                       3: //System 3
                           IF #_id_decoded_OP[#i].Device_Type = 30 THEN //VTD
                               "Screen_DB".OrderProcessing[#i] := CONCAT(IN1 := "System_DB_3".OrderTable[1].Device, IN2 := ' To LEVEL ', IN3 := #Level_Strg);
                           ELSIF #_id_decoded_OP[#i].Device_Type = 10 THEN //CNV1
                               "Screen_DB".OrderProcessing[#i] := CONCAT(IN1 := "System_DB_3".OrderTable[1].Device, IN2 := ' To CNV 1 LEVEL ', IN3 := #Level_Strg);
                           ELSIF #_id_decoded_OP[#i].Device_Type = 11 THEN //CNV2
                               "Screen_DB".OrderProcessing[#i] := CONCAT(IN1 := "System_DB_3".OrderTable[1].Device, IN2 := ' To CNV 2 LEVEL ', IN3 := #Level_Strg);
                           ELSIF #_id_decoded_OP[#i].Device_Type = 12 THEN //ECONVEYOR
                               "Screen_DB".OrderProcessing[#i] := CONCAT(IN1 := "System_DB_3".OrderTable[1].Device, IN2 := ' To ECONV LEVEL ', IN3 := #Level_Strg);
                           END_IF;

                       4: //System 4
                           IF #_id_decoded_OP[#i].Device_Type = 30 THEN //VTD
                               "Screen_DB".OrderProcessing[#i] := CONCAT(IN1 := "System_DB_4".OrderTable[1].Device, IN2 := ' To LEVEL ', IN3 := #Level_Strg);
                           ELSIF #_id_decoded_OP[#i].Device_Type = 10 THEN //CNV1
                               "Screen_DB".OrderProcessing[#i] := CONCAT(IN1 := "System_DB_4".OrderTable[1].Device, IN2 := ' To CNV 1 LEVEL ', IN3 := #Level_Strg);
                           ELSIF #_id_decoded_OP[#i].Device_Type = 11 THEN //CNV2
                               "Screen_DB".OrderProcessing[#i] := CONCAT(IN1 := "System_DB_4".OrderTable[1].Device, IN2 := ' To CNV 2 LEVEL ', IN3 := #Level_Strg);
                           ELSIF #_id_decoded_OP[#i].Device_Type = 12 THEN //ECONVEYOR
                               "Screen_DB".OrderProcessing[#i] := CONCAT(IN1 := "System_DB_4".OrderTable[1].Device, IN2 := ' To ECONV LEVEL ', IN3 := #Level_Strg);
                           END_IF;

                       5: //System 5
                           IF #_id_decoded_OP[#i].Device_Type = 30 THEN //VTD
                               "Screen_DB".OrderProcessing[#i] := CONCAT(IN1 := "System_DB_5".OrderTable[1].Device, IN2 := ' To LEVEL ', IN3 := #Level_Strg);
                           ELSIF #_id_decoded_OP[#i].Device_Type = 10 THEN //CNV1
                               "Screen_DB".OrderProcessing[#i] := CONCAT(IN1 := "System_DB_5".OrderTable[1].Device, IN2 := ' To CNV 1 LEVEL ', IN3 := #Level_Strg);
                           ELSIF #_id_decoded_OP[#i].Device_Type = 11 THEN //CNV2
                               "Screen_DB".OrderProcessing[#i] := CONCAT(IN1 := "System_DB_5".OrderTable[1].Device, IN2 := ' To CNV 2 LEVEL ', IN3 := #Level_Strg);
                           ELSIF #_id_decoded_OP[#i].Device_Type = 12 THEN //ECONVEYOR
                               "Screen_DB".OrderProcessing[#i] := CONCAT(IN1 := "System_DB_5".OrderTable[1].Device, IN2 := ' To ECONV LEVEL ', IN3 := #Level_Strg);
                           END_IF;
                   END_CASE;
               END_IF;
               END_FOR;

       END_REGION

       //empty background
       IF "System_DB_1".Error OR "System_DB_2".Error OR "System_DB_3".Error OR "System_DB_4".Error OR "System_DB_5".Error OR
           "Error_Word_1" <> 0 OR
           "Errors_Profinet_1" <> 0 OR
           "Errors_Profinet_2" <> 0 OR
           "Errors_Profinet_3" <> 0 OR
           "Errors_Profinet_4" <> 0 OR
           "Errors_Profinet_5" <> 0 OR
           "Errors_Profinet_6" <> 0 OR
           "Errors_Profinet_7" <> 0 OR
           "Errors_Profinet_8" <> 0 OR
           "Errors_Profinet_9" <> 0 OR
           "Errors_Profinet_10".%X0 OR
           "Errors_Profinet_10".%X1 OR
           "Errors_Profinet_10".%X2 OR
           "Errors_Profinet_10".%X3 OR
           "Errors_Profinet_10".%X4 OR
           "Errors_Profinet_10".%X5 OR
           "Errors_Profinet_10".%X6 OR
           "Errors_Profinet_10".%X7 OR
           "Errors_Profinet_10".%X8 OR
           "Errors_Profinet_10".%X9 OR
           "Errors_Profinet_10".%X10 OR
           "Errors_Profinet_10".%X11 OR
           "Errors_Profinet_10".%X12 OR
           "Errors_Profinet_10".%X13 OR
           "Errors_Profinet_11" <> 0 OR
           "Erros_Supply_Feedback_1" <> 0 OR
           "Erros_Supply_Feedback_2" <> 0 OR
           "Erros_Supply_Feedback_3" <> 0 OR
           "Erros_Supply_Feedback_4" <> 0 OR
           "Erros_Supply_Feedback_5" <> 0 OR
           "Erros_Supply_Feedback_6" <> 0 OR
           "Erros_Supply_Feedback_7" <> 0 OR
           "Sick Lector_Error code 1" <> 0 OR
           "Sick Lector_Error code 2" <> 0 OR
           "Sick Lector_Error code 3" <> 0 OR
           "Sick Lector_Error code 4" <> 0 OR
           "Sick Lector_Error code 5" <> 0 OR
           "Linear Encoder_Device Errors 1" <> 0 OR
           "Linear Encoder_Device Errors 2" <> 0 OR
           "Linear Encoder_Device Errors 3" <> 0 OR
           "Linear Encoder_Device Errors 4" <> 0 OR
           "Linear Encoder_Device Errors 5" <> 0 OR
           "Estop_Error_Word_1" <> 0 OR
           "Estop_Error_Word_2" <> 0 OR
           "Estop_Error_Word_3" <> 0 OR
           "Estop_Error_Word_4" <> 0 OR
           "Estop_Error_Word_5" <> 0 OR
           "Estop_Error_Word_6" <> 0 OR
           "Errors_Word_LightGuard_1" <> 0
       THEN
           "Screen_DB".EmptyTemplate_Background := 1;
       ELSE
           "Screen_DB".EmptyTemplate_Background := 0;
       END_IF;    //e

       // //main background - DEVICES
       // IF "HMI_DB".ScreenNo_Main = 1 AND "VTD_System_Selected_HMI" <> 0 THEN //VTD SCREEN
       //     IF "Control_DB".VTD_Sys["VTD_System_Selected_HMI"]."Error" THEN
       //         "Screen_DB".MainTemplate_Background := 1;
       //     ELSE
       //         "Screen_DB".MainTemplate_Background := 0;
       //     END_IF;
       // ELSIF "HMI_DB".ScreenNo_Main = 2 AND "CNV_System_Selected" <> 0 AND "CNV2_Selected" <> 0 AND "CNV_Level_Selected" <> 0 THEN //CONVEYOR SCREEN
       //     IF "CNV2_Selected" = 1 AND ("Control_DB".LCnv_Sys["CNV_System_Selected"].Cnv_Level["CNV_Level_Selected"].Cnv1.Error OR
       //         "Control_DB".ECnv_Sys["CNV_System_Selected"].Error) THEN
       //         "Screen_DB".MainTemplate_Background := 1;
       //     ELSIF "CNV2_Selected" = 2 AND ("Control_DB".LCnv_Sys["CNV_System_Selected"].Cnv_Level["CNV_Level_Selected"].Cnv2.Error OR
       //         "Control_DB".ECnv_Sys["CNV_System_Selected"].Error) THEN
       //         "Screen_DB".MainTemplate_Background := 1;
       //     ELSE
       //         "Screen_DB".MainTemplate_Background := 0;
       //     END_IF;
       // ELSE
       //     "Screen_DB".MainTemplate_Background := 0;
       // END_IF;
   END_REGION;

   REGION SHUTTLES
       IF "Screen_DB".Shuttle_Select >= 1 AND "Screen_DB".Shuttle_Select <= "Settings_DB".System.Shuttle_Count THEN
           CASE "Screen_DB".Shuttle_Select OF
               1:
                   "Screen_DB".Shuttle := "Shuttle_MQTT_DB".Shuttle_MQTT[1].Message.Shuttle_Status;
               2:
                   "Screen_DB".Shuttle := "Shuttle_MQTT_DB".Shuttle_MQTT[2].Message.Shuttle_Status;
               3:
                   "Screen_DB".Shuttle := "Shuttle_MQTT_DB".Shuttle_MQTT[3].Message.Shuttle_Status;
               4:
                   "Screen_DB".Shuttle := "Shuttle_MQTT_DB".Shuttle_MQTT[4].Message.Shuttle_Status;
               5:
                   "Screen_DB".Shuttle := "Shuttle_MQTT_DB".Shuttle_MQTT[5].Message.Shuttle_Status;
               6:
                   "Screen_DB".Shuttle := "Shuttle_MQTT_DB".Shuttle_MQTT[6].Message.Shuttle_Status;
               7:
                   "Screen_DB".Shuttle := "Shuttle_MQTT_DB".Shuttle_MQTT[7].Message.Shuttle_Status;
               8:
                   "Screen_DB".Shuttle := "Shuttle_MQTT_DB".Shuttle_MQTT[8].Message.Shuttle_Status;
               9:
                   "Screen_DB".Shuttle := "Shuttle_MQTT_DB".Shuttle_MQTT[9].Message.Shuttle_Status;
               10:
                   "Screen_DB".Shuttle := "Shuttle_MQTT_DB".Shuttle_MQTT[10].Message.Shuttle_Status;
               11:
                   "Screen_DB".Shuttle := "Shuttle_MQTT_DB".Shuttle_MQTT[11].Message.Shuttle_Status;
               12:
                   "Screen_DB".Shuttle := "Shuttle_MQTT_DB".Shuttle_MQTT[12].Message.Shuttle_Status;
               13:
                   "Screen_DB".Shuttle := "Shuttle_MQTT_DB".Shuttle_MQTT[13].Message.Shuttle_Status;
               14:
                   "Screen_DB".Shuttle := "Shuttle_MQTT_DB".Shuttle_MQTT[14].Message.Shuttle_Status;
               15:
                   "Screen_DB".Shuttle := "Shuttle_MQTT_DB".Shuttle_MQTT[15].Message.Shuttle_Status;
               16:
                   "Screen_DB".Shuttle := "Shuttle_MQTT_DB".Shuttle_MQTT[16].Message.Shuttle_Status;
               17:
                   "Screen_DB".Shuttle := "Shuttle_MQTT_DB".Shuttle_MQTT[17].Message.Shuttle_Status;
               18:
                   "Screen_DB".Shuttle := "Shuttle_MQTT_DB".Shuttle_MQTT[18].Message.Shuttle_Status;
               19:
                   "Screen_DB".Shuttle := "Shuttle_MQTT_DB".Shuttle_MQTT[19].Message.Shuttle_Status;
               20:
                   "Screen_DB".Shuttle := "Shuttle_MQTT_DB".Shuttle_MQTT[20].Message.Shuttle_Status;
               21:
                   "Screen_DB".Shuttle := "Shuttle_MQTT_DB".Shuttle_MQTT[21].Message.Shuttle_Status;
               22:
                   "Screen_DB".Shuttle := "Shuttle_MQTT_DB".Shuttle_MQTT[22].Message.Shuttle_Status;
               23:
                   "Screen_DB".Shuttle := "Shuttle_MQTT_DB".Shuttle_MQTT[23].Message.Shuttle_Status;
               // 24:
               //     "Screen_DB".Shuttle := "Shuttle_MQTT_DB".Shuttle_MQTT[24].Message.Shuttle_Status;
           END_CASE;
       END_IF;

       //E-STOP
       IF "Charge_Shuttle_Commands" THEN
           CASE "Shuttle_Level_Selected" OF
               1:
                   "Shuttle_Level_EStop" := "L1_Estop";
               2:
                   "Shuttle_Level_EStop" := "L2_Estop";
               3:
                   "Shuttle_Level_EStop" := "L3_Estop";
               4:
                   "Shuttle_Level_EStop" := "L4_Estop";
               5:
                   "Shuttle_Level_EStop" := "L5_Estop";
               6:
                   "Shuttle_Level_EStop" := "L6_Estop";
               7:
                   "Shuttle_Level_EStop" := "L7_Estop";
               8:
                   "Shuttle_Level_EStop" := "L8_Estop";
           END_CASE;
       ELSE
           CASE "Shuttle_Level_Selected" OF
               1:
                   "L1_Estop" := "Shuttle_Level_EStop";
               2:
                   "L2_Estop" := "Shuttle_Level_EStop";
               3:
                   "L3_Estop" := "Shuttle_Level_EStop";
               4:
                   "L4_Estop" := "Shuttle_Level_EStop";
               5:
                   "L5_Estop" := "Shuttle_Level_EStop";
               6:
                   "L6_Estop" := "Shuttle_Level_EStop";
               7:
                   "L7_Estop" := "Shuttle_Level_EStop";
               8:
                   "L8_Estop" := "Shuttle_Level_EStop";
           END_CASE;
       END_IF;
   END_REGION

   REGION ORDER TABLE
       //CHARGE OT DATA
       IF "Screen_DB".Charge_OT THEN
           CASE "Main_OrderTable_Selected" OF
               1:
                   "OT_Charge_Commands"("Auto_Test_1_DB");
               2:
                   "OT_Charge_Commands"("Auto_Test_2_DB");
               3:
                   "OT_Charge_Commands"("Auto_Test_3_DB");
               4:
                   "OT_Charge_Commands_1"("Auto_Test_4_DB");
               5:
                   "OT_Charge_Commands_1"("Auto_Test_5_DB");
           END_CASE;
           "T_Charge_OT".TON(IN := TRUE,
                             PT := T#1000ms);
           IF "T_Charge_OT".Q THEN
               "T_Charge_OT".TON(IN := FALSE,
                                 PT := T#0ms);
               "Screen_DB".Charge_OT := FALSE;
           END_IF;
       END_IF;

       IF NOT "Screen_DB".Charge_OT THEN
           "T_Charge_OT".TON(IN := FALSE,
                             PT := T#0ms);

           CASE "Main_OrderTable_Selected" OF
               1:
                   "Clear_OT(1)" := "Clear_OT";
                   "FC_Orders"(Sys := 1,
                               System := "System_DB_1",
                               Auto_Test := "Auto_Test_1_DB",
                               VTD_CurrentOrder := "Order_Table_FB_DB_1".VTD_CurrentOrder,
                               Pallet_InOut_CurrentOrder := "Order_Table_FB_DB_1".Pallet_InOut_CurrentOrder,
                               Shuttle_InOut_CurrentOrder := "Order_Table_FB_DB_1".Shuttle_InOut_CurrentOrder,
                               System_Busy := "System_1_Busy");

               2:
                   "Clear_OT(2)" := "Clear_OT";
                   "FC_Orders"(Sys := 2,
                               System := "System_DB_2",
                               Auto_Test := "Auto_Test_2_DB",
                               VTD_CurrentOrder := "Order_Table_FB_DB_2".VTD_CurrentOrder,
                               Pallet_InOut_CurrentOrder := "Order_Table_FB_DB_2".Pallet_InOut_CurrentOrder,
                               Shuttle_InOut_CurrentOrder := "Order_Table_FB_DB_2".Shuttle_InOut_CurrentOrder,
                               System_Busy := "System_2_Busy");

               3:
                   "Clear_OT(3)" := "Clear_OT";
                   "FC_Orders"(Sys := 3,
                               System := "System_DB_3",
                               Auto_Test := "Auto_Test_3_DB",
                               VTD_CurrentOrder := "Order_Table_FB_DB_3".VTD_CurrentOrder,
                               Pallet_InOut_CurrentOrder := "Order_Table_FB_DB_3".Pallet_InOut_CurrentOrder,
                               Shuttle_InOut_CurrentOrder := "Order_Table_FB_DB_3".Shuttle_InOut_CurrentOrder,
                               System_Busy := "System_3_Busy");

               4:
                   "Clear_OT(4)" := "Clear_OT";
                   "FC_Orders_2"(Sys := 4,
                               System := "System_DB_4",
                               Auto_Test := "Auto_Test_4_DB",
                               VTD_CurrentOrder := "Order_Table_FB_DB_4".VTD_CurrentOrder,
                               Pallet_InOut_CurrentOrder := "Order_Table_FB_DB_4".Pallet_InOut_CurrentOrder,
                               Shuttle_InOut_CurrentOrder := "Order_Table_FB_DB_4".Shuttle_InOut_CurrentOrder,
                               System_Busy := "System_4_Busy");

               5:
                   "Clear_OT(5)" := "Clear_OT";
                   "FC_Orders_2"(Sys := 5,
                               System := "System_DB_5",
                               Auto_Test := "Auto_Test_5_DB",
                               VTD_CurrentOrder := "Order_Table_FB_DB_5".VTD_CurrentOrder,
                               Pallet_InOut_CurrentOrder := "Order_Table_FB_DB_5".Pallet_InOut_CurrentOrder,
                               Shuttle_InOut_CurrentOrder := "Order_Table_FB_DB_5".Shuttle_InOut_CurrentOrder,
                               System_Busy := "System_5_Busy");

           END_CASE;
       END_IF;
   END_REGION

   "HMI_DB".Password := '12345';

   REGION VTD BARCODE
       CASE "VTD_System_Selected_HMI" OF
           1:
               "Screen_DB".VTD_Barcode := "Control_DB".VTDBarcode_Station[1].Barcode;
               "Screen_DB".VTD_Barcode_Visu := "Control_DB".VTDBarcode_Station[1].Barcode <> '';
           2:
               "Screen_DB".VTD_Barcode := "Control_DB".VTDBarcode_Station[2].Barcode;
               "Screen_DB".VTD_Barcode_Visu := "Control_DB".VTDBarcode_Station[2].Barcode <> '';
           3:
               "Screen_DB".VTD_Barcode := "Control_DB".VTDBarcode_Station[3].Barcode;
               "Screen_DB".VTD_Barcode_Visu := "Control_DB".VTDBarcode_Station[3].Barcode <> '';
           4:
               "Screen_DB".VTD_Barcode := "Control_DB".VTDBarcode_Station[4].Barcode;
               "Screen_DB".VTD_Barcode_Visu := "Control_DB".VTDBarcode_Station[4].Barcode <> '';
           5:
               "Screen_DB".VTD_Barcode := "Control_DB".VTDBarcode_Station[5].Barcode;
               "Screen_DB".VTD_Barcode_Visu := "Control_DB".VTDBarcode_Station[5].Barcode <> '';
       END_CASE;
   END_REGION VTD BARCODE

   // IF "FirstScan" THEN
       "TCPIP_Enable" := TRUE;
   // ELSE
       // "TCP_IP_Shuttle_DB_1".enable :=
       // "TCP_IP_Shuttle_DB_2".enable :=
       // "TCP_IP_Shuttle_DB_3".enable :=
       // "TCP_IP_Shuttle_DB_4".enable :=
       // "TCP_IP_Shuttle_DB_5".enable :=
       // "TCP_IP_Shuttle_DB_6".enable :=
       // "TCP_IP_Shuttle_DB_7".enable :=
       // "TCP_IP_Shuttle_DB_8".enable :=
       // "TCP_IP_Shuttle_DB_9".enable :=
       // "TCP_IP_Shuttle_DB_10".enable :=
       // "TCP_IP_Shuttle_DB_11".enable :=
       // "TCP_IP_Shuttle_DB_12".enable :=
       // "TCP_IP_Shuttle_DB_13".enable :=
       // "TCP_IP_Shuttle_DB_14".enable :=
       // "TCP_IP_Shuttle_DB_15".enable :=
       // "TCP_IP_Shuttle_DB_16".enable :=
       // "TCP_IP_Shuttle_DB_17".enable :=
       // "TCP_IP_Shuttle_DB_18".enable :=
       // "TCP_IP_Shuttle_DB_19".enable :=
       // "TCP_IP_Shuttle_DB_20".enable :=
       // "TCP_IP_Shuttle_DB_21".enable :=
       // "TCP_IP_Shuttle_DB_22".enable :=
       // "TCP_IP_Shuttle_DB_23".enable := "TCPIP_Enable";
   // END_IF;
END_FUNCTION

FUNCTION "Screens_2" : Void   // FC61, SCL
{ S7_Optimized_Access := 'TRUE' }
VERSION : 0.1
// stored: AutoNumber true, IsIECCheckEnabled false, SetENOAutomatically false, UDAEnableTagReadback false
   VAR_INPUT
      HMI_No : UInt;
      Sys_No : UInt;
   END_VAR
   VAR_TEMP
      i : UInt;
      j : UInt;
   END_VAR
BEGIN
   REGION MAIN SCREEN
       //main background - DEVICES
       IF "HMI_DB".ScreenNo[#HMI_No] = 1 THEN //VTD SCREEN
       //     IF "Control_DB".VTD_Sys["VTD_System_Selected_HMI"]."Error" THEN
       //         "Screen_DB_1".MainTemplate_Background := 1;
       //     ELSE
       //         "Screen_DB_1".MainTemplate_Background := 0;
       //     END_IF;
       // ELSIF "HMI_DB".ScreenNo = 2 AND "CNV_System_Selected" <> 0 AND "CNV2_Selected" <> 0 THEN //CONVEYOR SCREEN
       //     IF "CNV2_Selected" = 1 AND ("Control_DB".LCnv_Sys["CNV_System_Selected"].Cnv_Level["CNV_Level_Selected"].Cnv1.Error OR
       //         "Control_DB".ECnv_Sys["CNV_System_Selected"].Error) THEN
       //         "Screen_DB_1".MainTemplate_Background := 1;
       //     ELSIF "CNV2_Selected" = 2 AND ("Control_DB".LCnv_Sys["CNV_System_Selected"].Cnv_Level["CNV_Level_Selected"].Cnv2.Error OR
       //         "Control_DB".ECnv_Sys["CNV_System_Selected"].Error) THEN
       //         "Screen_DB_1".MainTemplate_Background := 1;
       //     ELSE
       //         "Screen_DB_1".MainTemplate_Background := 0;
       //     END_IF;
       //     
           ;
       ELSE
           "Screen_DB_1".MainTemplate_Background[#HMI_No] := 0;
       END_IF;
   END_REGION;

   REGION SHUTTLES
       CASE "Screen_DB_1".Shuttle_Select[#HMI_No] OF
           1:
               "Screen_DB_1".Shuttle := "Shuttle_MQTT_DB".Shuttle_MQTT[1].Message.Shuttle_Status;
           2:
               "Screen_DB_1".Shuttle := "Shuttle_MQTT_DB".Shuttle_MQTT[2].Message.Shuttle_Status;
           3:
               "Screen_DB_1".Shuttle := "Shuttle_MQTT_DB".Shuttle_MQTT[3].Message.Shuttle_Status;
           4:
               "Screen_DB_1".Shuttle := "Shuttle_MQTT_DB".Shuttle_MQTT[4].Message.Shuttle_Status;
           5:
               "Screen_DB_1".Shuttle := "Shuttle_MQTT_DB".Shuttle_MQTT[5].Message.Shuttle_Status;
           6:
               "Screen_DB_1".Shuttle := "Shuttle_MQTT_DB".Shuttle_MQTT[6].Message.Shuttle_Status;
           7:
               "Screen_DB_1".Shuttle := "Shuttle_MQTT_DB".Shuttle_MQTT[7].Message.Shuttle_Status;
           8:
               "Screen_DB_1".Shuttle := "Shuttle_MQTT_DB".Shuttle_MQTT[8].Message.Shuttle_Status;
           9:
               "Screen_DB_1".Shuttle := "Shuttle_MQTT_DB".Shuttle_MQTT[9].Message.Shuttle_Status;
           10:
               "Screen_DB_1".Shuttle := "Shuttle_MQTT_DB".Shuttle_MQTT[10].Message.Shuttle_Status;
           11:
               "Screen_DB_1".Shuttle := "Shuttle_MQTT_DB".Shuttle_MQTT[11].Message.Shuttle_Status;
           12:
               "Screen_DB_1".Shuttle := "Shuttle_MQTT_DB".Shuttle_MQTT[12].Message.Shuttle_Status;
           13:
               "Screen_DB_1".Shuttle := "Shuttle_MQTT_DB".Shuttle_MQTT[13].Message.Shuttle_Status;
           14:
               "Screen_DB_1".Shuttle := "Shuttle_MQTT_DB".Shuttle_MQTT[14].Message.Shuttle_Status;
           15:
               "Screen_DB_1".Shuttle := "Shuttle_MQTT_DB".Shuttle_MQTT[15].Message.Shuttle_Status;
           16:
               "Screen_DB_1".Shuttle := "Shuttle_MQTT_DB".Shuttle_MQTT[16].Message.Shuttle_Status;
           17:
               "Screen_DB_1".Shuttle := "Shuttle_MQTT_DB".Shuttle_MQTT[17].Message.Shuttle_Status;
           18:
               "Screen_DB_1".Shuttle := "Shuttle_MQTT_DB".Shuttle_MQTT[18].Message.Shuttle_Status;
           19:
               "Screen_DB_1".Shuttle := "Shuttle_MQTT_DB".Shuttle_MQTT[19].Message.Shuttle_Status;
           20:
               "Screen_DB_1".Shuttle := "Shuttle_MQTT_DB".Shuttle_MQTT[20].Message.Shuttle_Status;
           21:
               "Screen_DB_1".Shuttle := "Shuttle_MQTT_DB".Shuttle_MQTT[21].Message.Shuttle_Status;
           22:
               "Screen_DB_1".Shuttle := "Shuttle_MQTT_DB".Shuttle_MQTT[22].Message.Shuttle_Status;
           23:
               "Screen_DB_1".Shuttle := "Shuttle_MQTT_DB".Shuttle_MQTT[23].Message.Shuttle_Status;
       END_CASE;
   END_REGION

   REGION ORDER TABLE
           CASE #Sys_No OF
               1:
                   "Clear_OT(1)" := "Clear_OT";
                   "FC_Orders_1"(Sys := 1,
                               System := "System_DB_1",
                               VTD_CurrentOrder := "Order_Table_FB_DB_1".VTD_CurrentOrder,
                               Pallet_InOut_CurrentOrder := "Order_Table_FB_DB_1".Pallet_InOut_CurrentOrder,
                               Shuttle_InOut_CurrentOrder := "Order_Table_FB_DB_1".Shuttle_InOut_CurrentOrder);

               2:
                   "Clear_OT(2)" := "Clear_OT";
                   "FC_Orders_1"(Sys := 2,
                               System := "System_DB_2",
                               VTD_CurrentOrder := "Order_Table_FB_DB_2".VTD_CurrentOrder,
                               Pallet_InOut_CurrentOrder := "Order_Table_FB_DB_2".Pallet_InOut_CurrentOrder,
                               Shuttle_InOut_CurrentOrder := "Order_Table_FB_DB_2".Shuttle_InOut_CurrentOrder);

               3:
                   "Clear_OT(3)" := "Clear_OT";
                   "FC_Orders_1"(Sys := 3,
                               System := "System_DB_3",
                               VTD_CurrentOrder := "Order_Table_FB_DB_3".VTD_CurrentOrder,
                               Pallet_InOut_CurrentOrder := "Order_Table_FB_DB_3".Pallet_InOut_CurrentOrder,
                               Shuttle_InOut_CurrentOrder := "Order_Table_FB_DB_3".Shuttle_InOut_CurrentOrder);

               4:
                   "Clear_OT(4)" := "Clear_OT";
                   "FC_Orders_1"(Sys := 4,
                               System := "System_DB_4",
                               VTD_CurrentOrder := "Order_Table_FB_DB_4".VTD_CurrentOrder,
                               Pallet_InOut_CurrentOrder := "Order_Table_FB_DB_4".Pallet_InOut_CurrentOrder,
                               Shuttle_InOut_CurrentOrder := "Order_Table_FB_DB_4".Shuttle_InOut_CurrentOrder);

               5:
                   "Clear_OT(5)" := "Clear_OT";
                   "FC_Orders_1"(Sys := 5,
                               System := "System_DB_5",
                               VTD_CurrentOrder := "Order_Table_FB_DB_5".VTD_CurrentOrder,
                               Pallet_InOut_CurrentOrder := "Order_Table_FB_DB_5".Pallet_InOut_CurrentOrder,
                               Shuttle_InOut_CurrentOrder := "Order_Table_FB_DB_5".Shuttle_InOut_CurrentOrder);

           END_CASE;
   END_REGION

   REGION ALARMS
       //HMI 1
       IF "HMI_Box_Connected_1" = 6 OR ("HMI_Box_Connected_1" >= 11 AND "HMI_Box_Connected_1" <= 19) THEN
           IF "Screen_DB_1".Alarm_Current_Buttons[#HMI_No] THEN
               "Screen_DB_1".Alarms_ActiveTable[#HMI_No] := 1;
           ELSIF "Screen_DB_1".Alarm_History_Buttons[#HMI_No] THEN
               "Screen_DB_1".Alarms_ActiveTable[#HMI_No] := 11;
           END_IF;
       ELSIF "HMI_Box_Connected_1" >= 21 AND "HMI_Box_Connected_1" <= 29 THEN
           IF "Screen_DB_1".Alarm_Current_Buttons[#HMI_No] THEN
               "Screen_DB_1".Alarms_ActiveTable[#HMI_No] := 2;
           ELSIF "Screen_DB_1".Alarm_History_Buttons[#HMI_No] THEN
               "Screen_DB_1".Alarms_ActiveTable[#HMI_No] := 21;
           END_IF;
       ELSIF "HMI_Box_Connected_1" >= 31 AND "HMI_Box_Connected_1" <= 39 THEN
           IF "Screen_DB_1".Alarm_Current_Buttons[#HMI_No] THEN
               "Screen_DB_1".Alarms_ActiveTable[#HMI_No] := 3;
           ELSIF "Screen_DB_1".Alarm_History_Buttons[#HMI_No] THEN
               "Screen_DB_1".Alarms_ActiveTable[#HMI_No] := 31;
           END_IF;
       ELSIF "HMI_Box_Connected_1">= 41 AND"HMI_Box_Connected_1" <= 49 THEN
           IF "Screen_DB_1".Alarm_Current_Buttons[#HMI_No] THEN
               "Screen_DB_1".Alarms_ActiveTable[#HMI_No] := 4;
           ELSIF "Screen_DB_1".Alarm_History_Buttons[#HMI_No] THEN
               "Screen_DB_1".Alarms_ActiveTable[#HMI_No] := 41;
           END_IF;
       ELSIF "HMI_Box_Connected_1" >= 51 AND "HMI_Box_Connected_1" <= 59 THEN
           IF "Screen_DB_1".Alarm_Current_Buttons[#HMI_No] THEN
               "Screen_DB_1".Alarms_ActiveTable[#HMI_No] := 5;
           ELSIF "Screen_DB_1".Alarm_History_Buttons[#HMI_No] THEN
               "Screen_DB_1".Alarms_ActiveTable[#HMI_No] := 51;
           END_IF;
       END_IF;
   END_REGION ;
END_FUNCTION

FUNCTION "Set_Bit_F" : Void   // FC7, SCL
{ S7_Optimized_Access := 'TRUE' }
VERSION : 0.1
// stored: AutoNumber true, IsIECCheckEnabled false, SetENOAutomatically false, UDAEnableTagReadback false
   VAR_INPUT
      Bit : UInt;
      Bit_Value : Bool;
   END_VAR
   VAR_IN_OUT
      Var : Word;
   END_VAR
BEGIN
   IF #Bit_Value THEN
       // Set the bit
       #Var := #Var OR SHL(IN := WORD#1, N := #Bit);
   // ELSE
   //     // Reset the bit
   //     #Var := #Var OR SHL(IN := DWORD#1, N := #Bit);
   END_IF;
END_FUNCTION

FUNCTION "Settings_Limits_FC" : Void   // FC65, SCL
{ S7_Optimized_Access := 'TRUE' }
VERSION : 0.1
// stored: AutoNumber true, IsIECCheckEnabled false, SetENOAutomatically false, UDAEnableTagReadback false
   VAR_IN_OUT
      VTD_Settings : "VTD_Settings";
   END_VAR
BEGIN
   IF #VTD_Settings.Lowest_Level < 1 THEN
       #VTD_Settings.Lowest_Level := 1;
   END_IF;

   IF #VTD_Settings.Highest_Level > 8 THEN
       #VTD_Settings.Lowest_Level := 8;
   END_IF;

   IF #VTD_Settings.Creep_Speed < 3 THEN
       #VTD_Settings.Creep_Speed := 3;
   END_IF;

   IF #VTD_Settings.Slow_Speed < 3 THEN
       #VTD_Settings.Slow_Speed := 3;
   END_IF;

   IF #VTD_Settings.Loaded_Speed < #VTD_Settings.Slow_Calib_Speed * 1.8 THEN
       #VTD_Settings.Loaded_Speed := #VTD_Settings.Slow_Calib_Speed * 1.8;
   END_IF;

   IF #VTD_Settings.Shuttle_Speed < #VTD_Settings.Slow_Calib_Speed * 1.8 THEN
       #VTD_Settings.Shuttle_Speed := #VTD_Settings.Slow_Calib_Speed * 1.8;
   END_IF;

   IF #VTD_Settings.Pallet_Speed < #VTD_Settings.Slow_Calib_Speed * 1.8 THEN
       #VTD_Settings.Pallet_Speed := #VTD_Settings.Slow_Calib_Speed * 1.8;
   END_IF;

   IF #VTD_Settings.Empty_Speed < #VTD_Settings.Slow_Calib_Speed * 1.8 THEN
       #VTD_Settings.Empty_Speed := #VTD_Settings.Slow_Calib_Speed * 1.8;
   END_IF;

   IF #VTD_Settings.Dock_speed > 10 THEN
       #VTD_Settings.Dock_speed := 10;
   END_IF;

   IF #VTD_Settings.Empty_Speed > 120 THEN
       #VTD_Settings.Empty_Speed := 120;
   END_IF;

   IF #VTD_Settings.Pallet_Speed > 120 THEN
       #VTD_Settings.Pallet_Speed := 120;
   END_IF;

   IF #VTD_Settings.Chain_Slack_Timeout > 5000 THEN
       #VTD_Settings.Chain_Slack_Timeout := 5000;
   END_IF;

   IF #VTD_Settings.Acc_Range_1 < 60 THEN
       #VTD_Settings.Acc_Range_1 := 60;
   END_IF;

   IF #VTD_Settings.Acc_Range_2 < 60 THEN
       #VTD_Settings.Acc_Range_2 := 60;
   END_IF;

   IF #VTD_Settings.Acc_Range_3 < 60 THEN
       #VTD_Settings.Acc_Range_3 := 60;
   END_IF;

   IF #VTD_Settings.Acc_Range_1 > 100 THEN
       #VTD_Settings.Acc_Range_1 := 100;
   END_IF;

   IF #VTD_Settings.Acc_Range_2 > 100 THEN
       #VTD_Settings.Acc_Range_2 := 100;
   END_IF;

   IF #VTD_Settings.Acc_Range_3 > 100 THEN
       #VTD_Settings.Acc_Range_3 := 100;
   END_IF;
END_FUNCTION

FUNCTION "VTD_Charge_Settings" : Void   // FC41, SCL
{ S7_Optimized_Access := 'TRUE' }
VERSION : 0.1
// stored: AutoNumber true, IsIECCheckEnabled false, SetENOAutomatically false, UDAEnableTagReadback false
BEGIN
   //VTD SETTINGS
   CASE "VTD_System_Selected_HMI" OF
       1:
           "PopUps_DB".VTD_Settings := "Settings_DB".VTD_Sys[1];
       2:
           "PopUps_DB".VTD_Settings := "Settings_DB".VTD_Sys[2];
       3:
           "PopUps_DB".VTD_Settings := "Settings_DB".VTD_Sys[3];
       4:
           "PopUps_DB".VTD_Settings := "Settings_DB".VTD_Sys[4];
       5:
           "PopUps_DB".VTD_Settings := "Settings_DB".VTD_Sys[5];
   END_CASE;
END_FUNCTION

FUNCTION "VTD_Charge_Settings_1" : Void   // FC58, SCL
{ S7_Optimized_Access := 'TRUE' }
VERSION : 0.1
// stored: AutoNumber true, IsIECCheckEnabled false, SetENOAutomatically false, UDAEnableTagReadback false
   VAR_INPUT
      HMI_Box : UInt;
      Sys_No : UInt;
   END_VAR
BEGIN
   "PopUps_DB_1"."VTD_Settings"[#HMI_Box] := "Settings_DB".VTD_Sys[#Sys_No];
   "PopUps_DB_1"."Shuttle_MQTT_Settings" := "Settings_DB".Shuttle_MQTT;
END_FUNCTION

FUNCTION_BLOCK "VTD_HMI_FB"   // FB14, SCL
{ S7_Optimized_Access := 'TRUE' }
VERSION : 0.1
// stored: AutoNumber true, IsIECCheckEnabled false, IsRetainMemResEnabled false, MemoryReserve 100, SetENOAutomatically false, UDAEnableTagReadback false
   VAR
      T_Charge { S7_SetPoint := 'True'} : TON_TIME;
   END_VAR
BEGIN
   //CHARGE DATA CHANGING CONVEYORS ID
   IF "VTD_System_Selected_HMI" <> "VTD_ID_HMI_OLD" THEN
       "Screen_DB".Charge_VTD_Commands := TRUE;
       "VTD_ID_HMI_OLD" := "VTD_System_Selected_HMI";
   END_IF;

   //CHARGE ONCE THE COMMANDS STATUS
   IF "Screen_DB".Charge_VTD_Commands THEN
       CASE "VTD_System_Selected_HMI" OF
           1:
               "VTD_Mode_Change_HMI" := "Control_DB".VTD_Sys[1].Mode;
               "VTD_Enable_HMI" := "Control_DB".VTD_Sys[1].Instruction.Enable;
               "LE_Bypass" := "LE_Bypass(1)";
               "VTD_Stop_HMI" := "Control_DB".VTD_Sys[1].Instruction.Stop;
           2:
               "VTD_Mode_Change_HMI" := "Control_DB".VTD_Sys[2].Mode;
               "VTD_Enable_HMI" := "Control_DB".VTD_Sys[2].Instruction.Enable;
               "LE_Bypass" := "LE_Bypass(2)";
               "VTD_Stop_HMI" := "Control_DB".VTD_Sys[2].Instruction.Stop;
           3:
               "VTD_Mode_Change_HMI" := "Control_DB".VTD_Sys[3].Mode;
               "VTD_Enable_HMI" := "Control_DB".VTD_Sys[3].Instruction.Enable;
               "LE_Bypass" := "LE_Bypass(3)";
               "VTD_Stop_HMI" := "Control_DB".VTD_Sys[3].Instruction.Stop;
           4:
               "VTD_Mode_Change_HMI" := "Control_DB".VTD_Sys[4].Mode;
               "VTD_Enable_HMI" := "Control_DB".VTD_Sys[4].Instruction.Enable;
               "LE_Bypass" := "LE_Bypass(4)";
               "VTD_Stop_HMI" := "Control_DB".VTD_Sys[4].Instruction.Stop;
           5:
               "VTD_Mode_Change_HMI" := "Control_DB".VTD_Sys[5].Mode;
               "VTD_Enable_HMI" := "Control_DB".VTD_Sys[5].Instruction.Enable;
               "LE_Bypass" := "LE_Bypass(5)";
               "VTD_Stop_HMI" := "Control_DB".VTD_Sys[5].Instruction.Stop;
       END_CASE;

       #T_Charge.TON(IN := TRUE,
                     PT := T#500mS);
       IF #T_Charge.Q THEN
           #T_Charge.TON(IN := FALSE,
                         PT := T#0mS);
           "Screen_DB".Charge_VTD_Commands := 0;
       END_IF;

   // CHARGE DATA FROM HMI (AFTER CHARGE DATA)
   ELSIF "HMI_DB".ScreenNo_Main = 1 AND NOT "Screen_DB".Charge_VTD_Commands THEN
       CASE "VTD_System_Selected_HMI" OF
           1:
               "Feed_VTD_HMI_FC"(Sys_No := 1,
                                 Rem_Loc_Keys:= "HMI_DB".Rem_Loc_Keys[1].Level,
                                 Safety_OK := "Remote_Panel_DB_1".Safety_OK,
                                 BCD_Test_Ok_HMI := "SICK_Lector_DB_1".Test_OK,
                                 BCD_Error_HMI := "SICK_Lector_DB_1".Error,
                                 BCD_RdDone := "SICK_Lector_DB_1".RdDone,
                                 BCD_ReqDone := "SICK_Lector_DB_1".ReqDone,
                                 BCD_ReqBusy := "SICK_Lector_DB_1".ReqBusy,
                                 Start_InBarcodeStation := "Start_InBarcodeStation_HMI",
                                 Sick_Lector_Reseult := "SICK_Lector_DB_1".Barcode_Result,
                                 Level_Below_Extractor := "VTD_FB_DB_1".LevelBelowExtractor,
                                 Speed_mm_s := "VTD_FB_DB_1".VTDSpeed_mm_s,
                                 LE_Bypass := "LE_Bypass(1)",
                                 BCD_Start_Comm_Test_HMI := "BCD_Test_Comm_HMI(1)",
                                 BCD_Enable_Trigger_HMI := "BCD_Enable_Trigger_HMI(1)",
                                 BCD_Disable_Trigger_HMI := "BCD_Disable_Trigger_HMI(1)",
                                 BCD_Execute_Function := "SICK_Lector_Control_DB_1".Enable_Req,
                                 System_Busy => "System_1_Busy");

           2:
               "Feed_VTD_HMI_FC"(Sys_No := 2,
                                 Rem_Loc_Keys:="HMI_DB".Rem_Loc_Keys[2].Level,
                                 Safety_OK := "Remote_Panel_DB_2".Safety_OK,
                                 BCD_Test_Ok_HMI := "SICK_Lector_DB_2".Test_OK,
                                 BCD_Error_HMI := "SICK_Lector_DB_2".Error,
                                 BCD_RdDone := "SICK_Lector_DB_2".RdDone,
                                 BCD_ReqDone := "SICK_Lector_DB_2".ReqDone,
                                 BCD_ReqBusy := "SICK_Lector_DB_2".ReqBusy,
                                 Start_InBarcodeStation := "Start_InBarcodeStation_HMI",
                                 Sick_Lector_Reseult := "SICK_Lector_DB_2".Barcode_Result,
                                 Level_Below_Extractor := "VTD_FB_DB_2".LevelBelowExtractor,
                                 Speed_mm_s := "VTD_FB_DB_2".VTDSpeed_mm_s,
                                 LE_Bypass := "LE_Bypass(2)",
                                 BCD_Start_Comm_Test_HMI := "BCD_Test_Comm_HMI(2)",
                                 BCD_Enable_Trigger_HMI := "BCD_Enable_Trigger_HMI(2)",
                                 BCD_Disable_Trigger_HMI := "BCD_Disable_Trigger_HMI(2)",
                                 BCD_Execute_Function := "SICK_Lector_Control_DB_2".Enable_Req,
                                 System_Busy => "System_2_Busy");
           3:
               "Feed_VTD_HMI_FC"(Sys_No := 3,
                                 Rem_Loc_Keys:="HMI_DB".Rem_Loc_Keys[3].Level,
                                 Safety_OK := "Remote_Panel_DB_3".Safety_OK,
                                 BCD_Test_Ok_HMI := "SICK_Lector_DB_3".Test_OK,
                                 BCD_Error_HMI := "SICK_Lector_DB_3".Error,
                                 BCD_RdDone := "SICK_Lector_DB_3".RdDone,
                                 BCD_ReqDone := "SICK_Lector_DB_3".ReqDone,
                                 BCD_ReqBusy := "SICK_Lector_DB_3".ReqBusy,
                                 Start_InBarcodeStation := "Start_InBarcodeStation_HMI",
                                 Sick_Lector_Reseult := "SICK_Lector_DB_3".Barcode_Result,
                                 Level_Below_Extractor := "VTD_FB_DB_3".LevelBelowExtractor,
                                 Speed_mm_s := "VTD_FB_DB_3".VTDSpeed_mm_s,
                                 LE_Bypass := "LE_Bypass(3)",
                                 BCD_Start_Comm_Test_HMI := "BCD_Test_Comm_HMI(3)",
                                 BCD_Enable_Trigger_HMI := "BCD_Enable_Trigger_HMI(3)",
                                 BCD_Disable_Trigger_HMI := "BCD_Disable_Trigger_HMI(3)",
                                 BCD_Execute_Function := "SICK_Lector_Control_DB_3".Enable_Req,
                                 System_Busy => "System_3_Busy");
           4:
               "Feed_VTD_HMI_FC"(Sys_No := 4,
                                 Rem_Loc_Keys:="HMI_DB".Rem_Loc_Keys[4].Level,
                                 Safety_OK := "Remote_Panel_DB_4".Safety_OK,
                                 BCD_Test_Ok_HMI := "SICK_Lector_DB_4".Test_OK,
                                 BCD_Error_HMI := "SICK_Lector_DB_4".Error,
                                 BCD_RdDone := "SICK_Lector_DB_4".RdDone,
                                 BCD_ReqDone := "SICK_Lector_DB_4".ReqDone,
                                 BCD_ReqBusy := "SICK_Lector_DB_4".ReqBusy,
                                 Start_InBarcodeStation := "Start_InBarcodeStation_HMI",
                                 Sick_Lector_Reseult := "SICK_Lector_DB_4".Barcode_Result,
                                 Level_Below_Extractor := "VTD_FB_DB_4".LevelBelowExtractor,
                                 Speed_mm_s := "VTD_FB_DB_4".VTDSpeed_mm_s,
                                 LE_Bypass := "LE_Bypass(4)",
                                 BCD_Start_Comm_Test_HMI := "BCD_Test_Comm_HMI(4)",
                                 BCD_Enable_Trigger_HMI := "BCD_Enable_Trigger_HMI(4)",
                                 BCD_Disable_Trigger_HMI := "BCD_Disable_Trigger_HMI(4)",
                                 BCD_Execute_Function := "SICK_Lector_Control_DB_4".Enable_Req,
                                 System_Busy => "System_4_Busy");
           5:
               "Feed_VTD_HMI_FC"(Sys_No := 5,
                                 Rem_Loc_Keys:="HMI_DB".Rem_Loc_Keys[5].Level,
                                 Safety_OK := "Remote_Panel_DB_5".Safety_OK,
                                 BCD_Test_Ok_HMI := "SICK_Lector_DB_5".Test_OK,
                                 BCD_Error_HMI := "SICK_Lector_DB_5".Error,
                                 BCD_RdDone := "SICK_Lector_DB_5".RdDone,
                                 BCD_ReqDone := "SICK_Lector_DB_5".ReqDone,
                                 BCD_ReqBusy := "SICK_Lector_DB_5".ReqBusy,
                                 Start_InBarcodeStation := "Start_InBarcodeStation_HMI",
                                 Sick_Lector_Reseult := "SICK_Lector_DB_5".Barcode_Result,
                                 Level_Below_Extractor := "VTD_FB_DB_5".LevelBelowExtractor,
                                 Speed_mm_s := "VTD_FB_DB_5".VTDSpeed_mm_s,
                                 LE_Bypass := "LE_Bypass(5)",
                                 BCD_Start_Comm_Test_HMI := "BCD_Test_Comm_HMI(5)",
                                 BCD_Enable_Trigger_HMI := "BCD_Enable_Trigger_HMI(5)",
                                 BCD_Disable_Trigger_HMI := "BCD_Disable_Trigger_HMI(5)",
                                 BCD_Execute_Function := "SICK_Lector_Control_DB_5".Enable_Req,
                                 System_Busy => "System_5_Busy");
       END_CASE;
   END_IF;
END_FUNCTION_BLOCK

FUNCTION_BLOCK "VTD_HMI_FB_1"   // FB15, SCL
{ S7_Optimized_Access := 'TRUE' }
VERSION : 0.1
// stored: AutoNumber true, IsIECCheckEnabled false, IsRetainMemResEnabled false, MemoryReserve 100, SetENOAutomatically false, UDAEnableTagReadback false
   VAR_INPUT
      HMI_No : UInt;
      HMI_Box { ExternalAccessible := 'False'; ExternalVisible := 'False'; ExternalWritable := 'False'} : UInt;
      Sys_No : UInt;
   END_VAR
   VAR
      T_Charge { S7_SetPoint := 'True'} : TON_TIME;
      T_Charge_IN : Bool;
      Charged : Bool;
   END_VAR
BEGIN
   //CHARGE ONCE THE COMMANDS STATUS
   IF NOT #T_Charge.Q THEN
       CASE #Sys_No OF
           1:
               "VTD_HMI".Mode_Change[#HMI_No] := "Control_DB".VTD_Sys[1].Mode;
               "VTD_HMI".Enable[#HMI_No] := "Control_DB".VTD_Sys[1].Instruction.Enable;
               "PopUps_DB_1".Linear_Encoder[#HMI_No].LE_Bypass := "VTD_HMI".LE_Bypass[1];
               "VTD_HMI".Stop[#HMI_No] := "Control_DB".VTD_Sys[1].Instruction.Stop;
           2:
               "VTD_HMI".Mode_Change[#HMI_No] := "Control_DB".VTD_Sys[2].Mode;
               "VTD_HMI".Enable[#HMI_No] := "Control_DB".VTD_Sys[2].Instruction.Enable;
               "PopUps_DB_1".Linear_Encoder[#HMI_No].LE_Bypass := "VTD_HMI".LE_Bypass[2];
               "VTD_HMI".Stop[#HMI_No] := "Control_DB".VTD_Sys[2].Instruction.Stop;
           3:
               "VTD_HMI".Mode_Change[#HMI_No] := "Control_DB".VTD_Sys[3].Mode;
               "VTD_HMI".Enable[#HMI_No] := "Control_DB".VTD_Sys[3].Instruction.Enable;
               "PopUps_DB_1".Linear_Encoder[#HMI_No].LE_Bypass := "VTD_HMI".LE_Bypass[3];
               "VTD_HMI".Stop[#HMI_No] := "Control_DB".VTD_Sys[3].Instruction.Stop;
           4:
               "VTD_HMI".Mode_Change[#HMI_No] := "Control_DB".VTD_Sys[4].Mode;
               "VTD_HMI".Enable[#HMI_No] := "Control_DB".VTD_Sys[4].Instruction.Enable;
               "PopUps_DB_1".Linear_Encoder[#HMI_No].LE_Bypass := "VTD_HMI".LE_Bypass[4];
               "VTD_HMI".Stop[#HMI_No] := "Control_DB".VTD_Sys[4].Instruction.Stop;
           5:
               "VTD_HMI".Mode_Change[#HMI_No] := "Control_DB".VTD_Sys[5].Mode;
               "VTD_HMI".Enable[#HMI_No] := "Control_DB".VTD_Sys[5].Instruction.Enable;
               "PopUps_DB_1".Linear_Encoder[#HMI_No].LE_Bypass := "VTD_HMI".LE_Bypass[5];
               "VTD_HMI".Stop[#HMI_No] := "Control_DB".VTD_Sys[5].Instruction.Stop;
       END_CASE;
       #T_Charge_IN := TRUE;
   END_IF;

   #T_Charge.TON(IN := #T_Charge_IN,
                 PT := T#500mS);
   IF #T_Charge.Q THEN
       #Charged := TRUE;
   END_IF;

   // CHARGE DATA FROM HMI (AFTER CHARGE DATA)
   "Control_DB".VTD_Sys[#Sys_No].Instruction.Mode_Change := 1;
   IF #Charged THEN
       CASE #Sys_No OF
           1:
               "Feed_VTD_HMI_FC_1"(HMI_No := #HMI_No,
                                   HMI_Box:= #HMI_Box,
                                   Sys_No := #Sys_No,
                                   Safety_OK := "Remote_Panel_DB_1".Safety_OK,
                                   BCD_Test_Ok_HMI := "SICK_Lector_DB_1".Test_OK,
                                   BCD_Error_HMI := "SICK_Lector_DB_1".Error,
                                   BCD_RdDone := "SICK_Lector_DB_1".RdDone,
                                   BCD_ReqDone := "SICK_Lector_DB_1".ReqDone,
                                   BCD_ReqBusy := "SICK_Lector_DB_1".ReqBusy,
                                   Sick_Lector_Reseult := "SICK_Lector_DB_1".Barcode_Result,
                                   Level_Below_Extractor := "VTD_FB_DB_1".LevelBelowExtractor,
                                   Speed_mm_s := "VTD_FB_DB_1".VTDSpeed_mm_s,
                                   BCD_Start_Comm_Test_HMI := "BCD_Test_Comm_HMI(1)",
                                   BCD_Enable_Trigger_HMI := "BCD_Enable_Trigger_HMI(1)",
                                   BCD_Disable_Trigger_HMI := "BCD_Disable_Trigger_HMI(1)",
                                   BCD_Execute_Function := "SICK_Lector_Control_DB_1".Enable_Req);

           2:
               "Feed_VTD_HMI_FC_1"(HMI_No := #HMI_No,
                                   HMI_Box:= #HMI_Box,
                                   Sys_No := #Sys_No,
                                   Safety_OK := "Remote_Panel_DB_2".Safety_OK,
                                   BCD_Test_Ok_HMI := "SICK_Lector_DB_2".Test_OK,
                                   BCD_Error_HMI := "SICK_Lector_DB_2".Error,
                                   BCD_RdDone := "SICK_Lector_DB_2".RdDone,
                                   BCD_ReqDone := "SICK_Lector_DB_2".ReqDone,
                                   BCD_ReqBusy := "SICK_Lector_DB_2".ReqBusy,
                                   Sick_Lector_Reseult := "SICK_Lector_DB_2".Barcode_Result,
                                   Level_Below_Extractor := "VTD_FB_DB_2".LevelBelowExtractor,
                                   Speed_mm_s := "VTD_FB_DB_2".VTDSpeed_mm_s,
                                   BCD_Start_Comm_Test_HMI := "BCD_Test_Comm_HMI(2)",
                                   BCD_Enable_Trigger_HMI := "BCD_Enable_Trigger_HMI(2)",
                                   BCD_Disable_Trigger_HMI := "BCD_Disable_Trigger_HMI(2)",
                                   BCD_Execute_Function := "SICK_Lector_Control_DB_2".Enable_Req);
           3:
               "Feed_VTD_HMI_FC_1"(HMI_No := #HMI_No,
                                   HMI_Box:= #HMI_Box,
                                   Sys_No := #Sys_No,
                                   Safety_OK := "Remote_Panel_DB_3".Safety_OK,
                                   BCD_Test_Ok_HMI := "SICK_Lector_DB_3".Test_OK,
                                   BCD_Error_HMI := "SICK_Lector_DB_3".Error,
                                   BCD_RdDone := "SICK_Lector_DB_3".RdDone,
                                   BCD_ReqDone := "SICK_Lector_DB_3".ReqDone,
                                   BCD_ReqBusy := "SICK_Lector_DB_3".ReqBusy,
                                   Sick_Lector_Reseult := "SICK_Lector_DB_3".Barcode_Result,
                                   Level_Below_Extractor := "VTD_FB_DB_3".LevelBelowExtractor,
                                   Speed_mm_s := "VTD_FB_DB_3".VTDSpeed_mm_s,
                                   BCD_Start_Comm_Test_HMI := "BCD_Test_Comm_HMI(3)",
                                   BCD_Enable_Trigger_HMI := "BCD_Enable_Trigger_HMI(3)",
                                   BCD_Disable_Trigger_HMI := "BCD_Disable_Trigger_HMI(3)",
                                   BCD_Execute_Function := "SICK_Lector_Control_DB_3".Enable_Req);
           4:
               "Feed_VTD_HMI_FC_1"(HMI_No := #HMI_No,
                                   HMI_Box:= #HMI_Box,
                                   Sys_No := #Sys_No,
                                   Safety_OK := "Remote_Panel_DB_4".Safety_OK,
                                   BCD_Test_Ok_HMI := "SICK_Lector_DB_4".Test_OK,
                                   BCD_Error_HMI := "SICK_Lector_DB_4".Error,
                                   BCD_RdDone := "SICK_Lector_DB_4".RdDone,
                                   BCD_ReqDone := "SICK_Lector_DB_4".ReqDone,
                                   BCD_ReqBusy := "SICK_Lector_DB_4".ReqBusy,
                                   Sick_Lector_Reseult := "SICK_Lector_DB_4".Barcode_Result,
                                   Level_Below_Extractor := "VTD_FB_DB_4".LevelBelowExtractor,
                                   Speed_mm_s := "VTD_FB_DB_4".VTDSpeed_mm_s,
                                   BCD_Start_Comm_Test_HMI := "BCD_Test_Comm_HMI(4)",
                                   BCD_Enable_Trigger_HMI := "BCD_Enable_Trigger_HMI(4)",
                                   BCD_Disable_Trigger_HMI := "BCD_Disable_Trigger_HMI(4)",
                                   BCD_Execute_Function := "SICK_Lector_Control_DB_4".Enable_Req);
           5:
               "Feed_VTD_HMI_FC_1"(HMI_No := #HMI_No,
                                   HMI_Box:= #HMI_Box,
                                   Sys_No := #Sys_No,
                                   Safety_OK := "Remote_Panel_DB_5".Safety_OK,
                                   BCD_Test_Ok_HMI := "SICK_Lector_DB_5".Test_OK,
                                   BCD_Error_HMI := "SICK_Lector_DB_5".Error,
                                   BCD_RdDone := "SICK_Lector_DB_5".RdDone,
                                   BCD_ReqDone := "SICK_Lector_DB_5".ReqDone,
                                   BCD_ReqBusy := "SICK_Lector_DB_5".ReqBusy,
                                   Sick_Lector_Reseult := "SICK_Lector_DB_5".Barcode_Result,
                                   Level_Below_Extractor := "VTD_FB_DB_5".LevelBelowExtractor,
                                   Speed_mm_s := "VTD_FB_DB_5".VTDSpeed_mm_s,
                                   BCD_Start_Comm_Test_HMI := "BCD_Test_Comm_HMI(5)",
                                   BCD_Enable_Trigger_HMI := "BCD_Enable_Trigger_HMI(5)",
                                   BCD_Disable_Trigger_HMI := "BCD_Disable_Trigger_HMI(5)",
                                   BCD_Execute_Function := "SICK_Lector_Control_DB_5".Enable_Req);
       END_CASE;
   END_IF;
END_FUNCTION_BLOCK

FUNCTION "VTD_Order_FC" : Void   // FC45, SCL
{ S7_Optimized_Access := 'TRUE' }
VERSION : 0.1
// stored: AutoNumber true, IsIECCheckEnabled false, SetENOAutomatically false, UDAEnableTagReadback false
   VAR_INPUT
      i_Sys : UInt;
      Level : UInt;
   END_VAR
   VAR_IN_OUT
      StepTable_0 : "OrderTable_UDT";
   END_VAR
   VAR_TEMP
      StrSys : String;
      Concat1 : String;
      StrLev : String;
      Concat2 : String;
      ID : DInt;
   END_VAR
BEGIN
   #StrSys := UINT_TO_STRING(#i_Sys);
   // Remove "+"
   IF #StrSys[1] = '+' THEN
       #StrSys := RIGHT(IN := #StrSys, L := LEN(#StrSys) - 1);
   END_IF;

   #StrLev := UINT_TO_STRING(#Level);

   // Remove "+"
   IF #StrLev[1] = '+' THEN
       #StrLev := RIGHT(IN := #StrLev, L := LEN(#StrLev) - 1);
   END_IF;

   // Build ID
   #Concat1 := CONCAT(IN1 := '300', IN2 := #StrLev);
   #Concat2 := CONCAT(IN1 := #Concat1, IN2 := '0');
   #ID := STRING_TO_DINT(IN := CONCAT(IN1 := #Concat2, IN2 := #StrSys));

   "Feed_Steptable_FC"(CurrentTime := "Time".CurrentLocalTime,
                       Task_Type := 1,
                       Source_Location := 0,
                       Destination_Location := #ID,
                       Pallet_Type := 'C',
                       Pallet_Alignment := 'N',
                       Shuttle_ID:=0,
                       StepTable := #"StepTable_0");
END_FUNCTION

FUNCTION "VTD_Status_Update_FC" : Void   // FC48, SCL
{ S7_Optimized_Access := 'TRUE' }
VERSION : 0.1
// stored: AutoNumber true, IsIECCheckEnabled false, SetENOAutomatically false, UDAEnableTagReadback false
   VAR_INPUT
      Infeed_Auto_Mode : Bool;
      Infeed_Manual_Mode : Bool;
      Infeed_Maintenance : Bool;
      Infeed_Alarm : Bool;
      Infeed_Ready : Bool;
      Outfeed_Auto_Mode : Bool;
      Pallet_ID : Array[1..100] of Byte;
   END_VAR
   VAR_OUTPUT
      SM_To_LGX_VTD_Status : Byte;
   END_VAR
   VAR_IN_OUT
      Pallet_ID_Received : Bool;
   END_VAR
   VAR_TEMP
      tStatusByte : Byte;
      ArrayHasData : Bool;
      i : UInt;
   END_VAR
BEGIN
   #tStatusByte := 0;

       #tStatusByte.%X0 := #Infeed_Auto_Mode;
       #tStatusByte.%X1 := #Infeed_Manual_Mode;
       #tStatusByte.%X2 := #Infeed_Maintenance;
       #tStatusByte.%X3 := #Infeed_Ready;
       #tStatusByte.%X4 := #Infeed_Alarm;

       #ArrayHasData := FALSE;

       FOR #i := 1 TO 100 DO
           IF #Pallet_ID[#i] <> 0 THEN
               #ArrayHasData := TRUE;
               EXIT;
           END_IF;
       END_FOR;

       #tStatusByte.%X5 := #Pallet_ID_Received AND #ArrayHasData;
       #tStatusByte.%X6 := #Outfeed_Auto_Mode;

       IF #Pallet_ID_Received AND NOT #ArrayHasData THEN
           #Pallet_ID_Received := FALSE;
       END_IF;

       // Bit 5, 6: Free
       // 
       #SM_To_LGX_VTD_Status := #tStatusByte;
END_FUNCTION

DATA_BLOCK "Auto_Test_1_DB"   // DB4
VERSION : 0.1
// stored: AutoNumber true, DBAccessibleFromOPCUA true, InstanceOfName Auto_Test, InstanceOfType FB
"Auto_Test"
BEGIN
END_DATA_BLOCK

DATA_BLOCK "Auto_Test_2_DB"   // DB118
VERSION : 0.1
// stored: AutoNumber true, DBAccessibleFromOPCUA true, InstanceOfName Auto_Test, InstanceOfType FB
"Auto_Test"
BEGIN
END_DATA_BLOCK

DATA_BLOCK "Auto_Test_3_DB"   // DB117
VERSION : 0.1
// stored: AutoNumber true, DBAccessibleFromOPCUA true, InstanceOfName Auto_Test, InstanceOfType FB
"Auto_Test"
BEGIN
END_DATA_BLOCK

DATA_BLOCK "Auto_Test_4_DB"   // DB59
VERSION : 0.1
// stored: AutoNumber true, DBAccessibleFromOPCUA true, InstanceOfName Auto_Test_1, InstanceOfType FB
"Auto_Test_1"
BEGIN
END_DATA_BLOCK

DATA_BLOCK "Auto_Test_5_DB"   // DB435
VERSION : 0.1
// stored: AutoNumber true, DBAccessibleFromOPCUA true, InstanceOfName Auto_Test_1, InstanceOfType FB
"Auto_Test_1"
BEGIN
END_DATA_BLOCK

DATA_BLOCK "Auto_Test_DB"   // DB24
{ S7_Optimized_Access := 'TRUE' }
VERSION : 0.1
// stored: AutoNumber true, DBAccessibleFromOPCUA true, InstanceOfName Auto_Test_DB_UDT, InstanceOfType UDT, IsOnlyStoredInLoadMemory false, IsWriteProtectedInAS false
"Auto_Test_DB_UDT"
   // VAR
   //    System : Array[1..5] of "Auto_Test_UDT";
   // END_VAR
BEGIN
END_DATA_BLOCK

DATA_BLOCK "Barcode_FB_DB_1"   // DB144
VERSION : 0.1
// stored: AutoNumber true, DBAccessibleFromOPCUA true, InstanceOfName Barcode_Station_FB, InstanceOfType FB
"Barcode_Station_FB"
BEGIN
END_DATA_BLOCK

DATA_BLOCK "Barcode_FB_DB_2"   // DB331
VERSION : 0.1
// stored: AutoNumber true, DBAccessibleFromOPCUA true, InstanceOfName Barcode_Station_FB, InstanceOfType FB
"Barcode_Station_FB"
BEGIN
END_DATA_BLOCK

DATA_BLOCK "Barcode_FB_DB_3"   // DB330
VERSION : 0.1
// stored: AutoNumber true, DBAccessibleFromOPCUA true, InstanceOfName Barcode_Station_FB, InstanceOfType FB
"Barcode_Station_FB"
BEGIN
END_DATA_BLOCK

DATA_BLOCK "Barcode_FB_DB_4"   // DB328
VERSION : 0.1
// stored: AutoNumber true, DBAccessibleFromOPCUA true, InstanceOfName Barcode_Station_FB, InstanceOfType FB
"Barcode_Station_FB"
BEGIN
END_DATA_BLOCK

DATA_BLOCK "Barcode_FB_DB_5"   // DB329
VERSION : 0.1
// stored: AutoNumber true, DBAccessibleFromOPCUA true, InstanceOfName Barcode_Station_FB, InstanceOfType FB
"Barcode_Station_FB"
BEGIN
END_DATA_BLOCK

DATA_BLOCK "C1101_FB_DB"   // DB102
AUTHOR : Mertin Coetzee
VERSION : 0.1
// stored: AutoNumber true, DBAccessibleFromOPCUA true, InstanceOfName Buffer_Conveyor_FB, InstanceOfType FB
"Buffer_Conveyor_FB"
BEGIN
END_DATA_BLOCK

DATA_BLOCK "C1102_FB_DB"   // DB123
AUTHOR : Mertin Coetzee
VERSION : 0.1
// stored: AutoNumber true, DBAccessibleFromOPCUA true, InstanceOfName Buffer_Conveyor_FB, InstanceOfType FB
"Buffer_Conveyor_FB"
BEGIN
END_DATA_BLOCK

DATA_BLOCK "C1103_FB_DB"   // DB109
AUTHOR : Mertin Coetzee
VERSION : 0.1
// stored: AutoNumber true, DBAccessibleFromOPCUA true, InstanceOfName Buffer_Conveyor_FB, InstanceOfType FB
"Buffer_Conveyor_FB"
BEGIN
END_DATA_BLOCK

DATA_BLOCK "C1104_FB_DB"   // DB111
AUTHOR : Mertin Coetzee
VERSION : 0.1
// stored: AutoNumber true, DBAccessibleFromOPCUA true, InstanceOfName Buffer_Conveyor_FB, InstanceOfType FB
"Buffer_Conveyor_FB"
BEGIN
END_DATA_BLOCK

DATA_BLOCK "C1105_FB_DB"   // DB105
AUTHOR : Mertin Coetzee
VERSION : 0.1
// stored: AutoNumber true, DBAccessibleFromOPCUA true, InstanceOfName Buffer_Conveyor_FB, InstanceOfType FB
"Buffer_Conveyor_FB"
BEGIN
END_DATA_BLOCK

DATA_BLOCK "C1106_FB_DB"   // DB113
AUTHOR : Mertin Coetzee
VERSION : 0.1
// stored: AutoNumber true, DBAccessibleFromOPCUA true, InstanceOfName Buffer_Conveyor_FB, InstanceOfType FB
"Buffer_Conveyor_FB"
BEGIN
END_DATA_BLOCK

DATA_BLOCK "C1107_FB_DB"   // DB108
AUTHOR : Mertin Coetzee
VERSION : 0.1
// stored: AutoNumber true, DBAccessibleFromOPCUA true, InstanceOfName Buffer_Conveyor_FB, InstanceOfType FB
"Buffer_Conveyor_FB"
BEGIN
END_DATA_BLOCK

DATA_BLOCK "C1108_FB_DB"   // DB122
AUTHOR : Mertin Coetzee
VERSION : 0.1
// stored: AutoNumber true, DBAccessibleFromOPCUA true, InstanceOfName Buffer_Conveyor_FB, InstanceOfType FB
"Buffer_Conveyor_FB"
BEGIN
END_DATA_BLOCK

DATA_BLOCK "C1201_FB_DB"   // DB119
AUTHOR : Mertin Coetzee
VERSION : 0.1
// stored: AutoNumber true, DBAccessibleFromOPCUA true, InstanceOfName Buffer_Conveyor_FB, InstanceOfType FB
"Buffer_Conveyor_FB"
BEGIN
END_DATA_BLOCK

DATA_BLOCK "C1202_FB_DB"   // DB106
AUTHOR : Mertin Coetzee
VERSION : 0.1
// stored: AutoNumber true, DBAccessibleFromOPCUA true, InstanceOfName Buffer_Conveyor_FB, InstanceOfType FB
"Buffer_Conveyor_FB"
BEGIN
END_DATA_BLOCK

DATA_BLOCK "C1203_FB_DB"   // DB116
AUTHOR : Mertin Coetzee
VERSION : 0.1
// stored: AutoNumber true, DBAccessibleFromOPCUA true, InstanceOfName Buffer_Conveyor_FB, InstanceOfType FB
"Buffer_Conveyor_FB"
BEGIN
END_DATA_BLOCK

DATA_BLOCK "C1204_FB_DB"   // DB107
AUTHOR : Mertin Coetzee
VERSION : 0.1
// stored: AutoNumber true, DBAccessibleFromOPCUA true, InstanceOfName Buffer_Conveyor_FB, InstanceOfType FB
"Buffer_Conveyor_FB"
BEGIN
END_DATA_BLOCK

DATA_BLOCK "C1205_FB_DB"   // DB114
AUTHOR : Mertin Coetzee
VERSION : 0.1
// stored: AutoNumber true, DBAccessibleFromOPCUA true, InstanceOfName Buffer_Conveyor_FB, InstanceOfType FB
"Buffer_Conveyor_FB"
BEGIN
END_DATA_BLOCK

DATA_BLOCK "C1206_FB_DB"   // DB26
AUTHOR : Mertin Coetzee
VERSION : 0.1
// stored: AutoNumber true, DBAccessibleFromOPCUA true, InstanceOfName Buffer_Conveyor_FB, InstanceOfType FB
"Buffer_Conveyor_FB"
BEGIN
END_DATA_BLOCK

DATA_BLOCK "C1207_FB_DB"   // DB150
AUTHOR : Mertin Coetzee
VERSION : 0.1
// stored: AutoNumber true, DBAccessibleFromOPCUA true, InstanceOfName Buffer_Conveyor_FB, InstanceOfType FB
"Buffer_Conveyor_FB"
BEGIN
END_DATA_BLOCK

DATA_BLOCK "C1208_FB_DB"   // DB6
AUTHOR : Mertin Coetzee
VERSION : 0.1
// stored: AutoNumber true, DBAccessibleFromOPCUA true, InstanceOfName Buffer_Conveyor_FB, InstanceOfType FB
"Buffer_Conveyor_FB"
BEGIN
END_DATA_BLOCK

DATA_BLOCK "C2101_FB_DB"   // DB56
AUTHOR : Mertin Coetzee
VERSION : 0.1
// stored: AutoNumber true, DBAccessibleFromOPCUA true, InstanceOfName Buffer_Conveyor_FB, InstanceOfType FB
"Buffer_Conveyor_FB"
BEGIN
END_DATA_BLOCK

DATA_BLOCK "C2102_FB_DB"   // DB146
AUTHOR : Mertin Coetzee
VERSION : 0.1
// stored: AutoNumber true, DBAccessibleFromOPCUA true, InstanceOfName Buffer_Conveyor_FB, InstanceOfType FB
"Buffer_Conveyor_FB"
BEGIN
END_DATA_BLOCK

DATA_BLOCK "C2103_FB_DB"   // DB103
AUTHOR : Mertin Coetzee
VERSION : 0.1
// stored: AutoNumber true, DBAccessibleFromOPCUA true, InstanceOfName Buffer_Conveyor_FB, InstanceOfType FB
"Buffer_Conveyor_FB"
BEGIN
END_DATA_BLOCK

DATA_BLOCK "C2104_FB_DB"   // DB101
AUTHOR : Mertin Coetzee
VERSION : 0.1
// stored: AutoNumber true, DBAccessibleFromOPCUA true, InstanceOfName Buffer_Conveyor_FB, InstanceOfType FB
"Buffer_Conveyor_FB"
BEGIN
END_DATA_BLOCK

DATA_BLOCK "C2105_FB_DB"   // DB77
AUTHOR : Mertin Coetzee
VERSION : 0.1
// stored: AutoNumber true, DBAccessibleFromOPCUA true, InstanceOfName Buffer_Conveyor_FB, InstanceOfType FB
"Buffer_Conveyor_FB"
BEGIN
END_DATA_BLOCK

DATA_BLOCK "C2106_FB_DB"   // DB148
AUTHOR : Mertin Coetzee
VERSION : 0.1
// stored: AutoNumber true, DBAccessibleFromOPCUA true, InstanceOfName Buffer_Conveyor_FB, InstanceOfType FB
"Buffer_Conveyor_FB"
BEGIN
END_DATA_BLOCK

DATA_BLOCK "C2107_FB_DB"   // DB104
AUTHOR : Mertin Coetzee
VERSION : 0.1
// stored: AutoNumber true, DBAccessibleFromOPCUA true, InstanceOfName Buffer_Conveyor_FB, InstanceOfType FB
"Buffer_Conveyor_FB"
BEGIN
END_DATA_BLOCK

DATA_BLOCK "C2108_FB_DB"   // DB68
AUTHOR : Mertin Coetzee
VERSION : 0.1
// stored: AutoNumber true, DBAccessibleFromOPCUA true, InstanceOfName Buffer_Conveyor_FB, InstanceOfType FB
"Buffer_Conveyor_FB"
BEGIN
END_DATA_BLOCK

DATA_BLOCK "C2201_FB_DB"   // DB28
AUTHOR : Mertin Coetzee
VERSION : 0.1
// stored: AutoNumber true, DBAccessibleFromOPCUA true, InstanceOfName Buffer_Conveyor_FB, InstanceOfType FB
"Buffer_Conveyor_FB"
BEGIN
END_DATA_BLOCK

DATA_BLOCK "C2202_FB_DB"   // DB72
AUTHOR : Mertin Coetzee
VERSION : 0.1
// stored: AutoNumber true, DBAccessibleFromOPCUA true, InstanceOfName Buffer_Conveyor_FB, InstanceOfType FB
"Buffer_Conveyor_FB"
BEGIN
END_DATA_BLOCK

DATA_BLOCK "C2203_FB_DB"   // DB70
AUTHOR : Mertin Coetzee
VERSION : 0.1
// stored: AutoNumber true, DBAccessibleFromOPCUA true, InstanceOfName Buffer_Conveyor_FB, InstanceOfType FB
"Buffer_Conveyor_FB"
BEGIN
END_DATA_BLOCK

DATA_BLOCK "C2204_FB_DB"   // DB27
AUTHOR : Mertin Coetzee
VERSION : 0.1
// stored: AutoNumber true, DBAccessibleFromOPCUA true, InstanceOfName Buffer_Conveyor_FB, InstanceOfType FB
"Buffer_Conveyor_FB"
BEGIN
END_DATA_BLOCK

DATA_BLOCK "C2205_FB_DB"   // DB149
AUTHOR : Mertin Coetzee
VERSION : 0.1
// stored: AutoNumber true, DBAccessibleFromOPCUA true, InstanceOfName Buffer_Conveyor_FB, InstanceOfType FB
"Buffer_Conveyor_FB"
BEGIN
END_DATA_BLOCK

DATA_BLOCK "C2206_FB_DB"   // DB147
AUTHOR : Mertin Coetzee
VERSION : 0.1
// stored: AutoNumber true, DBAccessibleFromOPCUA true, InstanceOfName Buffer_Conveyor_FB, InstanceOfType FB
"Buffer_Conveyor_FB"
BEGIN
END_DATA_BLOCK

DATA_BLOCK "C2207_FB_DB"   // DB29
AUTHOR : Mertin Coetzee
VERSION : 0.1
// stored: AutoNumber true, DBAccessibleFromOPCUA true, InstanceOfName Buffer_Conveyor_FB, InstanceOfType FB
"Buffer_Conveyor_FB"
BEGIN
END_DATA_BLOCK

DATA_BLOCK "C2208_FB_DB"   // DB78
AUTHOR : Mertin Coetzee
VERSION : 0.1
// stored: AutoNumber true, DBAccessibleFromOPCUA true, InstanceOfName Buffer_Conveyor_FB, InstanceOfType FB
"Buffer_Conveyor_FB"
BEGIN
END_DATA_BLOCK

DATA_BLOCK "C3101_FB_DB"   // DB86
AUTHOR : Mertin Coetzee
VERSION : 0.1
// stored: AutoNumber true, DBAccessibleFromOPCUA true, InstanceOfName Buffer_Conveyor_FB, InstanceOfType FB
"Buffer_Conveyor_FB"
BEGIN
END_DATA_BLOCK

DATA_BLOCK "C3102_FB_DB"   // DB87
AUTHOR : Mertin Coetzee
VERSION : 0.1
// stored: AutoNumber true, DBAccessibleFromOPCUA true, InstanceOfName Buffer_Conveyor_FB, InstanceOfType FB
"Buffer_Conveyor_FB"
BEGIN
END_DATA_BLOCK

DATA_BLOCK "C3103_FB_DB"   // DB91
AUTHOR : Mertin Coetzee
VERSION : 0.1
// stored: AutoNumber true, DBAccessibleFromOPCUA true, InstanceOfName Buffer_Conveyor_FB, InstanceOfType FB
"Buffer_Conveyor_FB"
BEGIN
END_DATA_BLOCK

DATA_BLOCK "C3104_FB_DB"   // DB90
AUTHOR : Mertin Coetzee
VERSION : 0.1
// stored: AutoNumber true, DBAccessibleFromOPCUA true, InstanceOfName Buffer_Conveyor_FB, InstanceOfType FB
"Buffer_Conveyor_FB"
BEGIN
END_DATA_BLOCK

DATA_BLOCK "C3105_FB_DB"   // DB93
AUTHOR : Mertin Coetzee
VERSION : 0.1
// stored: AutoNumber true, DBAccessibleFromOPCUA true, InstanceOfName Buffer_Conveyor_FB, InstanceOfType FB
"Buffer_Conveyor_FB"
BEGIN
END_DATA_BLOCK

DATA_BLOCK "C3106_FB_DB"   // DB80
AUTHOR : Mertin Coetzee
VERSION : 0.1
// stored: AutoNumber true, DBAccessibleFromOPCUA true, InstanceOfName Buffer_Conveyor_FB, InstanceOfType FB
"Buffer_Conveyor_FB"
BEGIN
END_DATA_BLOCK

DATA_BLOCK "C3107_FB_DB"   // DB84
AUTHOR : Mertin Coetzee
VERSION : 0.1
// stored: AutoNumber true, DBAccessibleFromOPCUA true, InstanceOfName Buffer_Conveyor_FB, InstanceOfType FB
"Buffer_Conveyor_FB"
BEGIN
END_DATA_BLOCK

DATA_BLOCK "C3108_FB_DB"   // DB92
AUTHOR : Mertin Coetzee
VERSION : 0.1
// stored: AutoNumber true, DBAccessibleFromOPCUA true, InstanceOfName Buffer_Conveyor_FB, InstanceOfType FB
"Buffer_Conveyor_FB"
BEGIN
END_DATA_BLOCK

DATA_BLOCK "C3201_FB_DB"   // DB89
AUTHOR : Mertin Coetzee
VERSION : 0.1
// stored: AutoNumber true, DBAccessibleFromOPCUA true, InstanceOfName Buffer_Conveyor_FB, InstanceOfType FB
"Buffer_Conveyor_FB"
BEGIN
END_DATA_BLOCK

DATA_BLOCK "C3202_FB_DB"   // DB82
AUTHOR : Mertin Coetzee
VERSION : 0.1
// stored: AutoNumber true, DBAccessibleFromOPCUA true, InstanceOfName Buffer_Conveyor_FB, InstanceOfType FB
"Buffer_Conveyor_FB"
BEGIN
END_DATA_BLOCK

DATA_BLOCK "C3203_FB_DB"   // DB85
AUTHOR : Mertin Coetzee
VERSION : 0.1
// stored: AutoNumber true, DBAccessibleFromOPCUA true, InstanceOfName Buffer_Conveyor_FB, InstanceOfType FB
"Buffer_Conveyor_FB"
BEGIN
END_DATA_BLOCK

DATA_BLOCK "C3204_FB_DB"   // DB88
AUTHOR : Mertin Coetzee
VERSION : 0.1
// stored: AutoNumber true, DBAccessibleFromOPCUA true, InstanceOfName Buffer_Conveyor_FB, InstanceOfType FB
"Buffer_Conveyor_FB"
BEGIN
END_DATA_BLOCK

DATA_BLOCK "C3205_FB_DB"   // DB94
AUTHOR : Mertin Coetzee
VERSION : 0.1
// stored: AutoNumber true, DBAccessibleFromOPCUA true, InstanceOfName Buffer_Conveyor_FB, InstanceOfType FB
"Buffer_Conveyor_FB"
BEGIN
END_DATA_BLOCK

DATA_BLOCK "C3206_FB_DB"   // DB83
AUTHOR : Mertin Coetzee
VERSION : 0.1
// stored: AutoNumber true, DBAccessibleFromOPCUA true, InstanceOfName Buffer_Conveyor_FB, InstanceOfType FB
"Buffer_Conveyor_FB"
BEGIN
END_DATA_BLOCK

DATA_BLOCK "C3207_FB_DB"   // DB95
AUTHOR : Mertin Coetzee
VERSION : 0.1
// stored: AutoNumber true, DBAccessibleFromOPCUA true, InstanceOfName Buffer_Conveyor_FB, InstanceOfType FB
"Buffer_Conveyor_FB"
BEGIN
END_DATA_BLOCK

DATA_BLOCK "C3208_FB_DB"   // DB81
AUTHOR : Mertin Coetzee
VERSION : 0.1
// stored: AutoNumber true, DBAccessibleFromOPCUA true, InstanceOfName Buffer_Conveyor_FB, InstanceOfType FB
"Buffer_Conveyor_FB"
BEGIN
END_DATA_BLOCK

DATA_BLOCK "C4101_FB_DB"   // DB100
AUTHOR : Mertin Coetzee
VERSION : 0.1
// stored: AutoNumber true, DBAccessibleFromOPCUA true, InstanceOfName Buffer_Conveyor_FB, InstanceOfType FB
"Buffer_Conveyor_FB"
BEGIN
END_DATA_BLOCK

DATA_BLOCK "C4102_FB_DB"   // DB112
AUTHOR : Mertin Coetzee
VERSION : 0.1
// stored: AutoNumber true, DBAccessibleFromOPCUA true, InstanceOfName Buffer_Conveyor_FB, InstanceOfType FB
"Buffer_Conveyor_FB"
BEGIN
END_DATA_BLOCK

DATA_BLOCK "C4103_FB_DB"   // DB33
AUTHOR : Mertin Coetzee
VERSION : 0.1
// stored: AutoNumber true, DBAccessibleFromOPCUA true, InstanceOfName Buffer_Conveyor_FB, InstanceOfType FB
"Buffer_Conveyor_FB"
BEGIN
END_DATA_BLOCK

DATA_BLOCK "C4104_FB_DB"   // DB145
AUTHOR : Mertin Coetzee
VERSION : 0.1
// stored: AutoNumber true, DBAccessibleFromOPCUA true, InstanceOfName Buffer_Conveyor_FB, InstanceOfType FB
"Buffer_Conveyor_FB"
BEGIN
END_DATA_BLOCK

DATA_BLOCK "C4105_FB_DB"   // DB140
AUTHOR : Mertin Coetzee
VERSION : 0.1
// stored: AutoNumber true, DBAccessibleFromOPCUA true, InstanceOfName Buffer_Conveyor_FB, InstanceOfType FB
"Buffer_Conveyor_FB"
BEGIN
END_DATA_BLOCK

DATA_BLOCK "C4106_FB_DB"   // DB142
AUTHOR : Mertin Coetzee
VERSION : 0.1
// stored: AutoNumber true, DBAccessibleFromOPCUA true, InstanceOfName Buffer_Conveyor_FB, InstanceOfType FB
"Buffer_Conveyor_FB"
BEGIN
END_DATA_BLOCK

DATA_BLOCK "C4107_FB_DB"   // DB151
AUTHOR : Mertin Coetzee
VERSION : 0.1
// stored: AutoNumber true, DBAccessibleFromOPCUA true, InstanceOfName Buffer_Conveyor_FB, InstanceOfType FB
"Buffer_Conveyor_FB"
BEGIN
END_DATA_BLOCK

DATA_BLOCK "C4108_FB_DB"   // DB143
AUTHOR : Mertin Coetzee
VERSION : 0.1
// stored: AutoNumber true, DBAccessibleFromOPCUA true, InstanceOfName Buffer_Conveyor_FB, InstanceOfType FB
"Buffer_Conveyor_FB"
BEGIN
END_DATA_BLOCK

DATA_BLOCK "C5101_FB_DB"   // DB127
AUTHOR : Mertin Coetzee
VERSION : 0.1
// stored: AutoNumber true, DBAccessibleFromOPCUA true, InstanceOfName Buffer_Conveyor_FB, InstanceOfType FB
"Buffer_Conveyor_FB"
BEGIN
END_DATA_BLOCK

DATA_BLOCK "C5102_FB_DB"   // DB133
AUTHOR : Mertin Coetzee
VERSION : 0.1
// stored: AutoNumber true, DBAccessibleFromOPCUA true, InstanceOfName Buffer_Conveyor_FB, InstanceOfType FB
"Buffer_Conveyor_FB"
BEGIN
END_DATA_BLOCK

DATA_BLOCK "C5103_FB_DB"   // DB129
AUTHOR : Mertin Coetzee
VERSION : 0.1
// stored: AutoNumber true, DBAccessibleFromOPCUA true, InstanceOfName Buffer_Conveyor_FB, InstanceOfType FB
"Buffer_Conveyor_FB"
BEGIN
END_DATA_BLOCK

DATA_BLOCK "C5104_FB_DB"   // DB125
AUTHOR : Mertin Coetzee
VERSION : 0.1
// stored: AutoNumber true, DBAccessibleFromOPCUA true, InstanceOfName Buffer_Conveyor_FB, InstanceOfType FB
"Buffer_Conveyor_FB"
BEGIN
END_DATA_BLOCK

DATA_BLOCK "C5105_FB_DB"   // DB138
AUTHOR : Mertin Coetzee
VERSION : 0.1
// stored: AutoNumber true, DBAccessibleFromOPCUA true, InstanceOfName Buffer_Conveyor_FB, InstanceOfType FB
"Buffer_Conveyor_FB"
BEGIN
END_DATA_BLOCK

DATA_BLOCK "C5106_FB_DB"   // DB126
AUTHOR : Mertin Coetzee
VERSION : 0.1
// stored: AutoNumber true, DBAccessibleFromOPCUA true, InstanceOfName Buffer_Conveyor_FB, InstanceOfType FB
"Buffer_Conveyor_FB"
BEGIN
END_DATA_BLOCK

DATA_BLOCK "C5107_FB_DB"   // DB124
AUTHOR : Mertin Coetzee
VERSION : 0.1
// stored: AutoNumber true, DBAccessibleFromOPCUA true, InstanceOfName Buffer_Conveyor_FB, InstanceOfType FB
"Buffer_Conveyor_FB"
BEGIN
END_DATA_BLOCK

DATA_BLOCK "C5108_FB_DB"   // DB130
AUTHOR : Mertin Coetzee
VERSION : 0.1
// stored: AutoNumber true, DBAccessibleFromOPCUA true, InstanceOfName Buffer_Conveyor_FB, InstanceOfType FB
"Buffer_Conveyor_FB"
BEGIN
END_DATA_BLOCK

DATA_BLOCK "Conveyor_HMI_FB_1_DB"   // DB50
VERSION : 0.1
// stored: AutoNumber true, DBAccessibleFromOPCUA true, InstanceOfName Conveyor_HMI_FB_1, InstanceOfType FB
"Conveyor_HMI_FB_1"
BEGIN
END_DATA_BLOCK

DATA_BLOCK "Conveyor_HMI_FB_2_DB"   // DB61
VERSION : 0.1
// stored: AutoNumber true, DBAccessibleFromOPCUA true, InstanceOfName Conveyor_HMI_FB_1, InstanceOfType FB
"Conveyor_HMI_FB_1"
BEGIN
END_DATA_BLOCK

DATA_BLOCK "Conveyor_HMI_FB_DB"   // DB73
VERSION : 0.1
// stored: AutoNumber true, DBAccessibleFromOPCUA true, InstanceOfName Conveyor_HMI_FB, InstanceOfType FB
"Conveyor_HMI_FB"
BEGIN
END_DATA_BLOCK

DATA_BLOCK "Default_SupervisionDB"   // DB2
VERSION : 0.1
// stored: AutoNumber true, DBAccessibleFromOPCUA true, InstanceOfName Default_SupervisionFB, InstanceOfType FB
"Default_SupervisionFB"
   // VAR
   //    PC_Flags { ExternalWritable := 'False'; S7_SetPoint := 'True'} : PC_Flags_V2;
   //    State { ExternalWritable := 'False'; S7_SetPoint := 'True'} : SV_FB_State_V2;
   // END_VAR
BEGIN
END_DATA_BLOCK

DATA_BLOCK "ECnv_FB_DB_1"   // DB14
AUTHOR : Mertin Coetzee
VERSION : 0.1
// stored: AutoNumber true, DBAccessibleFromOPCUA true, InstanceOfName EConveyor_FB, InstanceOfType FB
"EConveyor_FB"
   // VAR_INPUT
   //    Id : UInt;
   //    Safety_OK_Delayed : Bool;
   //    Safety_OK : Bool;
   //    Cnv_Settings : "ECnv_Settings";
   //    VTD_Current_Level : UInt;
   //    CNV_In_Out : Bool;
   //    CNV1_2_Selected : UInt;
   // END_VAR
   // VAR_IN_OUT
   //    Cnv_Control : "ECnv_Control";
   //    SinaSpeed : SinaSpeed;
   // END_VAR
   // VAR
   //    State : UInt;
   //    Timer_Transfer { S7_SetPoint := 'True'} : TON_TIME;
   //    Watchdog { S7_SetPoint := 'True'} : TON_TIME;
   //    Transfer_Direction { S7_SetPoint := 'True'} : String;
   //    MainSetpoint : Int;
   //    SinaSpeed_Instance { S7_SetPoint := 'True'} : SinaSpeed;
   //    IEC_Timer_0_Instance_1 { S7_SetPoint := 'True'} : TON_TIME;
   //    R_TRIG_Instance { S7_SetPoint := 'True'} : R_TRIG;
   //    R_Start_DB { S7_SetPoint := 'True'} : R_TRIG;
   //    R_Stop_DB { S7_SetPoint := 'True'} : R_TRIG;
   //    ID_Decoded_From { S7_SetPoint := 'True'} : "ID_Decoded";
   //    ID_Decoded_To { S7_SetPoint := 'True'} : "ID_Decoded";
   //    R_Slow { S7_SetPoint := 'True'} : R_TRIG;
   //    T_Ramp { S7_SetPoint := 'True'} : TON_TIME;
   //    T_Ramp_In : Bool;
   //    VTD_Level : UInt;
   //    TCheck_PalletType { S7_SetPoint := 'True'} : TON_TIME;
   // END_VAR
BEGIN
END_DATA_BLOCK

DATA_BLOCK "ECnv_FB_DB_2"   // DB13
AUTHOR : Mertin Coetzee
VERSION : 0.1
// stored: AutoNumber true, DBAccessibleFromOPCUA true, InstanceOfName EConveyor_FB, InstanceOfType FB
"EConveyor_FB"
   // VAR_INPUT
   //    Id : UInt;
   //    Safety_OK_Delayed : Bool;
   //    Safety_OK : Bool;
   //    Cnv_Settings : "ECnv_Settings";
   //    VTD_Current_Level : UInt;
   //    CNV_In_Out : Bool;
   //    CNV1_2_Selected : UInt;
   // END_VAR
   // VAR_IN_OUT
   //    Cnv_Control : "ECnv_Control";
   //    SinaSpeed : SinaSpeed;
   // END_VAR
   // VAR
   //    State : UInt;
   //    Timer_Transfer { S7_SetPoint := 'True'} : TON_TIME;
   //    Watchdog { S7_SetPoint := 'True'} : TON_TIME;
   //    Transfer_Direction { S7_SetPoint := 'True'} : String;
   //    MainSetpoint : Int;
   //    SinaSpeed_Instance { S7_SetPoint := 'True'} : SinaSpeed;
   //    IEC_Timer_0_Instance_1 { S7_SetPoint := 'True'} : TON_TIME;
   //    R_TRIG_Instance { S7_SetPoint := 'True'} : R_TRIG;
   //    R_Start_DB { S7_SetPoint := 'True'} : R_TRIG;
   //    R_Stop_DB { S7_SetPoint := 'True'} : R_TRIG;
   //    ID_Decoded_From { S7_SetPoint := 'True'} : "ID_Decoded";
   //    ID_Decoded_To { S7_SetPoint := 'True'} : "ID_Decoded";
   //    R_Slow { S7_SetPoint := 'True'} : R_TRIG;
   //    T_Ramp { S7_SetPoint := 'True'} : TON_TIME;
   //    T_Ramp_In : Bool;
   //    VTD_Level : UInt;
   //    TCheck_PalletType { S7_SetPoint := 'True'} : TON_TIME;
   // END_VAR
BEGIN
END_DATA_BLOCK

DATA_BLOCK "ECnv_FB_DB_3"   // DB15
AUTHOR : Mertin Coetzee
VERSION : 0.1
// stored: AutoNumber true, DBAccessibleFromOPCUA true, InstanceOfName EConveyor_FB, InstanceOfType FB
"EConveyor_FB"
   // VAR_INPUT
   //    Id : UInt;
   //    Safety_OK_Delayed : Bool;
   //    Safety_OK : Bool;
   //    Cnv_Settings : "ECnv_Settings";
   //    VTD_Current_Level : UInt;
   //    CNV_In_Out : Bool;
   //    CNV1_2_Selected : UInt;
   // END_VAR
   // VAR_IN_OUT
   //    Cnv_Control : "ECnv_Control";
   //    SinaSpeed : SinaSpeed;
   // END_VAR
   // VAR
   //    State : UInt;
   //    Timer_Transfer { S7_SetPoint := 'True'} : TON_TIME;
   //    Watchdog { S7_SetPoint := 'True'} : TON_TIME;
   //    Transfer_Direction { S7_SetPoint := 'True'} : String;
   //    MainSetpoint : Int;
   //    SinaSpeed_Instance { S7_SetPoint := 'True'} : SinaSpeed;
   //    IEC_Timer_0_Instance_1 { S7_SetPoint := 'True'} : TON_TIME;
   //    R_TRIG_Instance { S7_SetPoint := 'True'} : R_TRIG;
   //    R_Start_DB { S7_SetPoint := 'True'} : R_TRIG;
   //    R_Stop_DB { S7_SetPoint := 'True'} : R_TRIG;
   //    ID_Decoded_From { S7_SetPoint := 'True'} : "ID_Decoded";
   //    ID_Decoded_To { S7_SetPoint := 'True'} : "ID_Decoded";
   //    R_Slow { S7_SetPoint := 'True'} : R_TRIG;
   //    T_Ramp { S7_SetPoint := 'True'} : TON_TIME;
   //    T_Ramp_In : Bool;
   //    VTD_Level : UInt;
   //    TCheck_PalletType { S7_SetPoint := 'True'} : TON_TIME;
   // END_VAR
BEGIN
END_DATA_BLOCK

DATA_BLOCK "ECnv_FB_DB_4"   // DB16
AUTHOR : Mertin Coetzee
VERSION : 0.1
// stored: AutoNumber true, DBAccessibleFromOPCUA true, InstanceOfName EConveyor_FB, InstanceOfType FB
"EConveyor_FB"
   // VAR_INPUT
   //    Id : UInt;
   //    Safety_OK_Delayed : Bool;
   //    Safety_OK : Bool;
   //    Cnv_Settings : "ECnv_Settings";
   //    VTD_Current_Level : UInt;
   //    CNV_In_Out : Bool;
   //    CNV1_2_Selected : UInt;
   // END_VAR
   // VAR_IN_OUT
   //    Cnv_Control : "ECnv_Control";
   //    SinaSpeed : SinaSpeed;
   // END_VAR
   // VAR
   //    State : UInt;
   //    Timer_Transfer { S7_SetPoint := 'True'} : TON_TIME;
   //    Watchdog { S7_SetPoint := 'True'} : TON_TIME;
   //    Transfer_Direction { S7_SetPoint := 'True'} : String;
   //    MainSetpoint : Int;
   //    SinaSpeed_Instance { S7_SetPoint := 'True'} : SinaSpeed;
   //    IEC_Timer_0_Instance_1 { S7_SetPoint := 'True'} : TON_TIME;
   //    R_TRIG_Instance { S7_SetPoint := 'True'} : R_TRIG;
   //    R_Start_DB { S7_SetPoint := 'True'} : R_TRIG;
   //    R_Stop_DB { S7_SetPoint := 'True'} : R_TRIG;
   //    ID_Decoded_From { S7_SetPoint := 'True'} : "ID_Decoded";
   //    ID_Decoded_To { S7_SetPoint := 'True'} : "ID_Decoded";
   //    R_Slow { S7_SetPoint := 'True'} : R_TRIG;
   //    T_Ramp { S7_SetPoint := 'True'} : TON_TIME;
   //    T_Ramp_In : Bool;
   //    VTD_Level : UInt;
   //    TCheck_PalletType { S7_SetPoint := 'True'} : TON_TIME;
   // END_VAR
BEGIN
END_DATA_BLOCK

DATA_BLOCK "ECnv_FB_DB_5"   // DB5
AUTHOR : Mertin Coetzee
VERSION : 0.1
// stored: AutoNumber true, DBAccessibleFromOPCUA true, InstanceOfName EConveyor_FB, InstanceOfType FB
"EConveyor_FB"
   // VAR_INPUT
   //    Id : UInt;
   //    Safety_OK_Delayed : Bool;
   //    Safety_OK : Bool;
   //    Cnv_Settings : "ECnv_Settings";
   //    VTD_Current_Level : UInt;
   //    CNV_In_Out : Bool;
   //    CNV1_2_Selected : UInt;
   // END_VAR
   // VAR_IN_OUT
   //    Cnv_Control : "ECnv_Control";
   //    SinaSpeed : SinaSpeed;
   // END_VAR
   // VAR
   //    State : UInt;
   //    Timer_Transfer { S7_SetPoint := 'True'} : TON_TIME;
   //    Watchdog { S7_SetPoint := 'True'} : TON_TIME;
   //    Transfer_Direction { S7_SetPoint := 'True'} : String;
   //    MainSetpoint : Int;
   //    SinaSpeed_Instance { S7_SetPoint := 'True'} : SinaSpeed;
   //    IEC_Timer_0_Instance_1 { S7_SetPoint := 'True'} : TON_TIME;
   //    R_TRIG_Instance { S7_SetPoint := 'True'} : R_TRIG;
   //    R_Start_DB { S7_SetPoint := 'True'} : R_TRIG;
   //    R_Stop_DB { S7_SetPoint := 'True'} : R_TRIG;
   //    ID_Decoded_From { S7_SetPoint := 'True'} : "ID_Decoded";
   //    ID_Decoded_To { S7_SetPoint := 'True'} : "ID_Decoded";
   //    R_Slow { S7_SetPoint := 'True'} : R_TRIG;
   //    T_Ramp { S7_SetPoint := 'True'} : TON_TIME;
   //    T_Ramp_In : Bool;
   //    VTD_Level : UInt;
   //    TCheck_PalletType { S7_SetPoint := 'True'} : TON_TIME;
   // END_VAR
BEGIN
END_DATA_BLOCK

DATA_BLOCK "FB_HeartBeat_DB"   // DB136
VERSION : 0.1
// stored: AutoNumber true, DBAccessibleFromOPCUA true, InstanceOfName FB_HeartBeat, InstanceOfType FB
"FB_HeartBeat"
BEGIN
   TimeOut.PT := T#10S;
   TimeOut.IN := TRUE;
   "Timer".PT := T#500MS;
   "Timer".IN := TRUE;
END_DATA_BLOCK

DATA_BLOCK "F_Lock_FB_DB_1"   // DB411, F_DB
VERSION : 0.1
// stored: AutoNumber true, DBAccessibleFromOPCUA true, InstanceOfName F_Lock_FB, InstanceOfType FB
"F_Lock_FB"
BEGIN
END_DATA_BLOCK

DATA_BLOCK "F_Lock_FB_DB_10"   // DB422, F_DB
VERSION : 0.1
// stored: AutoNumber true, DBAccessibleFromOPCUA true, InstanceOfName F_Lock_FB, InstanceOfType FB
"F_Lock_FB"
BEGIN
END_DATA_BLOCK

DATA_BLOCK "F_Lock_FB_DB_11"   // DB423, F_DB
VERSION : 0.1
// stored: AutoNumber true, DBAccessibleFromOPCUA true, InstanceOfName F_Lock_FB, InstanceOfType FB
"F_Lock_FB"
BEGIN
END_DATA_BLOCK

DATA_BLOCK "F_Lock_FB_DB_12"   // DB424, F_DB
VERSION : 0.1
// stored: AutoNumber true, DBAccessibleFromOPCUA true, InstanceOfName F_Lock_FB, InstanceOfType FB
"F_Lock_FB"
BEGIN
END_DATA_BLOCK

DATA_BLOCK "F_Lock_FB_DB_2"   // DB412, F_DB
VERSION : 0.1
// stored: AutoNumber true, DBAccessibleFromOPCUA true, InstanceOfName F_Lock_FB, InstanceOfType FB
"F_Lock_FB"
BEGIN
END_DATA_BLOCK

DATA_BLOCK "F_Lock_FB_DB_3"   // DB416, F_DB
VERSION : 0.1
// stored: AutoNumber true, DBAccessibleFromOPCUA true, InstanceOfName F_Lock_FB, InstanceOfType FB
"F_Lock_FB"
BEGIN
END_DATA_BLOCK

DATA_BLOCK "F_Lock_FB_DB_4"   // DB417, F_DB
VERSION : 0.1
// stored: AutoNumber true, DBAccessibleFromOPCUA true, InstanceOfName F_Lock_FB, InstanceOfType FB
"F_Lock_FB"
BEGIN
END_DATA_BLOCK

DATA_BLOCK "F_Lock_FB_DB_5"   // DB418, F_DB
VERSION : 0.1
// stored: AutoNumber true, DBAccessibleFromOPCUA true, InstanceOfName F_Lock_FB, InstanceOfType FB
"F_Lock_FB"
BEGIN
END_DATA_BLOCK

DATA_BLOCK "F_Lock_FB_DB_6"   // DB419, F_DB
VERSION : 0.1
// stored: AutoNumber true, DBAccessibleFromOPCUA true, InstanceOfName F_Lock_FB, InstanceOfType FB
"F_Lock_FB"
BEGIN
END_DATA_BLOCK

DATA_BLOCK "F_Lock_FB_DB_7"   // DB420, F_DB
VERSION : 0.1
// stored: AutoNumber true, DBAccessibleFromOPCUA true, InstanceOfName F_Lock_FB, InstanceOfType FB
"F_Lock_FB"
BEGIN
END_DATA_BLOCK

DATA_BLOCK "F_Lock_FB_DB_8"   // DB421, F_DB
VERSION : 0.1
// stored: AutoNumber true, DBAccessibleFromOPCUA true, InstanceOfName F_Lock_FB, InstanceOfType FB
"F_Lock_FB"
BEGIN
END_DATA_BLOCK

DATA_BLOCK "F_Lock_FB_DB_9"   // DB415, F_DB
VERSION : 0.1
// stored: AutoNumber true, DBAccessibleFromOPCUA true, InstanceOfName F_Lock_FB, InstanceOfType FB
"F_Lock_FB"
BEGIN
END_DATA_BLOCK

DATA_BLOCK "GateAccess_Station_FB_DB_1"   // DB425
VERSION : 0.1
// stored: AutoNumber true, DBAccessibleFromOPCUA true, InstanceOfName GateAccess_Station_FB, InstanceOfType FB
"GateAccess_Station_FB"
BEGIN
END_DATA_BLOCK

DATA_BLOCK "GateAccess_Station_FB_DB_10"   // DB432
VERSION : 0.1
// stored: AutoNumber true, DBAccessibleFromOPCUA true, InstanceOfName GateAccess_Station_FB, InstanceOfType FB
"GateAccess_Station_FB"
BEGIN
END_DATA_BLOCK

DATA_BLOCK "GateAccess_Station_FB_DB_11"   // DB433
VERSION : 0.1
// stored: AutoNumber true, DBAccessibleFromOPCUA true, InstanceOfName GateAccess_Station_FB, InstanceOfType FB
"GateAccess_Station_FB"
BEGIN
END_DATA_BLOCK

DATA_BLOCK "GateAccess_Station_FB_DB_12"   // DB434
VERSION : 0.1
// stored: AutoNumber true, DBAccessibleFromOPCUA true, InstanceOfName GateAccess_Station_FB, InstanceOfType FB
"GateAccess_Station_FB"
BEGIN
END_DATA_BLOCK

DATA_BLOCK "GateAccess_Station_FB_DB_2"   // DB426
VERSION : 0.1
// stored: AutoNumber true, DBAccessibleFromOPCUA true, InstanceOfName GateAccess_Station_FB, InstanceOfType FB
"GateAccess_Station_FB"
BEGIN
END_DATA_BLOCK

DATA_BLOCK "GateAccess_Station_FB_DB_3"   // DB427
VERSION : 0.1
// stored: AutoNumber true, DBAccessibleFromOPCUA true, InstanceOfName GateAccess_Station_FB, InstanceOfType FB
"GateAccess_Station_FB"
BEGIN
END_DATA_BLOCK

DATA_BLOCK "GateAccess_Station_FB_DB_4"   // DB428
VERSION : 0.1
// stored: AutoNumber true, DBAccessibleFromOPCUA true, InstanceOfName GateAccess_Station_FB, InstanceOfType FB
"GateAccess_Station_FB"
BEGIN
END_DATA_BLOCK

DATA_BLOCK "GateAccess_Station_FB_DB_5"   // DB429
VERSION : 0.1
// stored: AutoNumber true, DBAccessibleFromOPCUA true, InstanceOfName GateAccess_Station_FB, InstanceOfType FB
"GateAccess_Station_FB"
BEGIN
END_DATA_BLOCK

DATA_BLOCK "GateAccess_Station_FB_DB_6"   // DB430
VERSION : 0.1
// stored: AutoNumber true, DBAccessibleFromOPCUA true, InstanceOfName GateAccess_Station_FB, InstanceOfType FB
"GateAccess_Station_FB"
BEGIN
END_DATA_BLOCK

DATA_BLOCK "GateAccess_Station_FB_DB_7"   // DB431
VERSION : 0.1
// stored: AutoNumber true, DBAccessibleFromOPCUA true, InstanceOfName GateAccess_Station_FB, InstanceOfType FB
"GateAccess_Station_FB"
BEGIN
END_DATA_BLOCK

DATA_BLOCK "GateAccess_Station_FB_DB_8"   // DB414
VERSION : 0.1
// stored: AutoNumber true, DBAccessibleFromOPCUA true, InstanceOfName GateAccess_Station_FB, InstanceOfType FB
"GateAccess_Station_FB"
BEGIN
END_DATA_BLOCK

DATA_BLOCK "GateAccess_Station_FB_DB_9"   // DB413
VERSION : 0.1
// stored: AutoNumber true, DBAccessibleFromOPCUA true, InstanceOfName GateAccess_Station_FB, InstanceOfType FB
"GateAccess_Station_FB"
BEGIN
END_DATA_BLOCK

DATA_BLOCK "LCom_Comm_Shuttle_FB_DB_1"   // DB65
AUTHOR : APC_ERLF
FAMILY : LCom
VERSION : 2.1
// stored: AutoNumber true, DBAccessibleFromOPCUA true, InstanceOfName LCom_Communication_FB, InstanceOfType FB
"LCom_Communication_FB"
BEGIN
END_DATA_BLOCK

DATA_BLOCK "LCom_Comm_Shuttle_FB_DB_10"   // DB359
AUTHOR : APC_ERLF
FAMILY : LCom
VERSION : 2.1
// stored: AutoNumber true, DBAccessibleFromOPCUA true, InstanceOfName LCom_Communication_FB, InstanceOfType FB
"LCom_Communication_FB"
BEGIN
END_DATA_BLOCK

DATA_BLOCK "LCom_Comm_Shuttle_FB_DB_11"   // DB358
AUTHOR : APC_ERLF
FAMILY : LCom
VERSION : 2.1
// stored: AutoNumber true, DBAccessibleFromOPCUA true, InstanceOfName LCom_Communication_FB, InstanceOfType FB
"LCom_Communication_FB"
BEGIN
END_DATA_BLOCK

DATA_BLOCK "LCom_Comm_Shuttle_FB_DB_12"   // DB371
AUTHOR : APC_ERLF
FAMILY : LCom
VERSION : 2.1
// stored: AutoNumber true, DBAccessibleFromOPCUA true, InstanceOfName LCom_Communication_FB, InstanceOfType FB
"LCom_Communication_FB"
BEGIN
END_DATA_BLOCK

DATA_BLOCK "LCom_Comm_Shuttle_FB_DB_13"   // DB356
AUTHOR : APC_ERLF
FAMILY : LCom
VERSION : 2.1
// stored: AutoNumber true, DBAccessibleFromOPCUA true, InstanceOfName LCom_Communication_FB, InstanceOfType FB
"LCom_Communication_FB"
BEGIN
END_DATA_BLOCK

DATA_BLOCK "LCom_Comm_Shuttle_FB_DB_14"   // DB354
AUTHOR : APC_ERLF
FAMILY : LCom
VERSION : 2.1
// stored: AutoNumber true, DBAccessibleFromOPCUA true, InstanceOfName LCom_Communication_FB, InstanceOfType FB
"LCom_Communication_FB"
BEGIN
END_DATA_BLOCK

DATA_BLOCK "LCom_Comm_Shuttle_FB_DB_15"   // DB373
AUTHOR : APC_ERLF
FAMILY : LCom
VERSION : 2.1
// stored: AutoNumber true, DBAccessibleFromOPCUA true, InstanceOfName LCom_Communication_FB, InstanceOfType FB
"LCom_Communication_FB"
BEGIN
END_DATA_BLOCK

DATA_BLOCK "LCom_Comm_Shuttle_FB_DB_16"   // DB351
AUTHOR : APC_ERLF
FAMILY : LCom
VERSION : 2.1
// stored: AutoNumber true, DBAccessibleFromOPCUA true, InstanceOfName LCom_Communication_FB, InstanceOfType FB
"LCom_Communication_FB"
BEGIN
END_DATA_BLOCK

DATA_BLOCK "LCom_Comm_Shuttle_FB_DB_17"   // DB352
AUTHOR : APC_ERLF
FAMILY : LCom
VERSION : 2.1
// stored: AutoNumber true, DBAccessibleFromOPCUA true, InstanceOfName LCom_Communication_FB, InstanceOfType FB
"LCom_Communication_FB"
BEGIN
END_DATA_BLOCK

DATA_BLOCK "LCom_Comm_Shuttle_FB_DB_18"   // DB353
AUTHOR : APC_ERLF
FAMILY : LCom
VERSION : 2.1
// stored: AutoNumber true, DBAccessibleFromOPCUA true, InstanceOfName LCom_Communication_FB, InstanceOfType FB
"LCom_Communication_FB"
BEGIN
END_DATA_BLOCK

DATA_BLOCK "LCom_Comm_Shuttle_FB_DB_19"   // DB368
AUTHOR : APC_ERLF
FAMILY : LCom
VERSION : 2.1
// stored: AutoNumber true, DBAccessibleFromOPCUA true, InstanceOfName LCom_Communication_FB, InstanceOfType FB
"LCom_Communication_FB"
BEGIN
END_DATA_BLOCK

DATA_BLOCK "LCom_Comm_Shuttle_FB_DB_2"   // DB370
AUTHOR : APC_ERLF
FAMILY : LCom
VERSION : 2.1
// stored: AutoNumber true, DBAccessibleFromOPCUA true, InstanceOfName LCom_Communication_FB, InstanceOfType FB
"LCom_Communication_FB"
BEGIN
END_DATA_BLOCK

DATA_BLOCK "LCom_Comm_Shuttle_FB_DB_20"   // DB372
AUTHOR : APC_ERLF
FAMILY : LCom
VERSION : 2.1
// stored: AutoNumber true, DBAccessibleFromOPCUA true, InstanceOfName LCom_Communication_FB, InstanceOfType FB
"LCom_Communication_FB"
BEGIN
END_DATA_BLOCK

DATA_BLOCK "LCom_Comm_Shuttle_FB_DB_21"   // DB369
AUTHOR : APC_ERLF
FAMILY : LCom
VERSION : 2.1
// stored: AutoNumber true, DBAccessibleFromOPCUA true, InstanceOfName LCom_Communication_FB, InstanceOfType FB
"LCom_Communication_FB"
BEGIN
END_DATA_BLOCK

DATA_BLOCK "LCom_Comm_Shuttle_FB_DB_22"   // DB365
AUTHOR : APC_ERLF
FAMILY : LCom
VERSION : 2.1
// stored: AutoNumber true, DBAccessibleFromOPCUA true, InstanceOfName LCom_Communication_FB, InstanceOfType FB
"LCom_Communication_FB"
BEGIN
END_DATA_BLOCK

DATA_BLOCK "LCom_Comm_Shuttle_FB_DB_23"   // DB366
AUTHOR : APC_ERLF
FAMILY : LCom
VERSION : 2.1
// stored: AutoNumber true, DBAccessibleFromOPCUA true, InstanceOfName LCom_Communication_FB, InstanceOfType FB
"LCom_Communication_FB"
BEGIN
END_DATA_BLOCK

DATA_BLOCK "LCom_Comm_Shuttle_FB_DB_24"   // DB355
AUTHOR : APC_ERLF
FAMILY : LCom
VERSION : 2.1
// stored: AutoNumber true, DBAccessibleFromOPCUA true, InstanceOfName LCom_Communication_FB, InstanceOfType FB
"LCom_Communication_FB"
BEGIN
END_DATA_BLOCK

DATA_BLOCK "LCom_Comm_Shuttle_FB_DB_3"   // DB357
AUTHOR : APC_ERLF
FAMILY : LCom
VERSION : 2.1
// stored: AutoNumber true, DBAccessibleFromOPCUA true, InstanceOfName LCom_Communication_FB, InstanceOfType FB
"LCom_Communication_FB"
BEGIN
END_DATA_BLOCK

DATA_BLOCK "LCom_Comm_Shuttle_FB_DB_4"   // DB367
AUTHOR : APC_ERLF
FAMILY : LCom
VERSION : 2.1
// stored: AutoNumber true, DBAccessibleFromOPCUA true, InstanceOfName LCom_Communication_FB, InstanceOfType FB
"LCom_Communication_FB"
BEGIN
END_DATA_BLOCK

DATA_BLOCK "LCom_Comm_Shuttle_FB_DB_5"   // DB364
AUTHOR : APC_ERLF
FAMILY : LCom
VERSION : 2.1
// stored: AutoNumber true, DBAccessibleFromOPCUA true, InstanceOfName LCom_Communication_FB, InstanceOfType FB
"LCom_Communication_FB"
BEGIN
END_DATA_BLOCK

DATA_BLOCK "LCom_Comm_Shuttle_FB_DB_6"   // DB363
AUTHOR : APC_ERLF
FAMILY : LCom
VERSION : 2.1
// stored: AutoNumber true, DBAccessibleFromOPCUA true, InstanceOfName LCom_Communication_FB, InstanceOfType FB
"LCom_Communication_FB"
BEGIN
END_DATA_BLOCK

DATA_BLOCK "LCom_Comm_Shuttle_FB_DB_7"   // DB362
AUTHOR : APC_ERLF
FAMILY : LCom
VERSION : 2.1
// stored: AutoNumber true, DBAccessibleFromOPCUA true, InstanceOfName LCom_Communication_FB, InstanceOfType FB
"LCom_Communication_FB"
BEGIN
END_DATA_BLOCK

DATA_BLOCK "LCom_Comm_Shuttle_FB_DB_8"   // DB361
AUTHOR : APC_ERLF
FAMILY : LCom
VERSION : 2.1
// stored: AutoNumber true, DBAccessibleFromOPCUA true, InstanceOfName LCom_Communication_FB, InstanceOfType FB
"LCom_Communication_FB"
BEGIN
END_DATA_BLOCK

DATA_BLOCK "LCom_Comm_Shuttle_FB_DB_9"   // DB360
AUTHOR : APC_ERLF
FAMILY : LCom
VERSION : 2.1
// stored: AutoNumber true, DBAccessibleFromOPCUA true, InstanceOfName LCom_Communication_FB, InstanceOfType FB
"LCom_Communication_FB"
BEGIN
END_DATA_BLOCK

DATA_BLOCK "LMQTT_Client_DB"   // DB158
AUTHOR : Siemens Industry Online Support
FAMILY : LMQTT
VERSION : 4.0
// stored: AutoNumber true, DBAccessibleFromOPCUA true, InstanceOfName LMQTT_Client, InstanceOfType FB
"LMQTT_Client"
BEGIN
END_DATA_BLOCK

DATA_BLOCK "LMQTT_Client_fb"   // DB42
AUTHOR : Siemens Industry Online Support
FAMILY : LMQTT
VERSION : 4.0
// stored: AutoNumber true, DBAccessibleFromOPCUA true, InstanceOfName LMQTT_Client, InstanceOfType FB
"LMQTT_Client"
BEGIN
END_DATA_BLOCK

DATA_BLOCK "LMQTT_DB"   // DB43
{ S7_Optimized_Access := 'TRUE' }
VERSION : 0.1
// stored: AutoNumber true, DBAccessibleFromOPCUA true, InstanceOfName LMQTT_DB_UDT, InstanceOfType UDT, IsOnlyStoredInLoadMemory false, IsWriteProtectedInAS false
"LMQTT_DB_UDT"
   // VAR
   //    enable : Bool;
   //    publish : Bool;
   //    subscribe : Bool;
   //    unsubscribe : Bool;
   //    qos : USInt;
   //    retain : Bool;
   //    publishMsgLen : UDInt;
   //    willMsgLen : UInt;
   //    connParam : "LMQTT_typeConnParam";
   //    clientIdentifier : WString;
   //    username : WString;
   //    password : WString;
   //    willtopic : WString;
   //    willMsgPayload : Array[1..128] of Byte;
   //    mqttTopic : WString;
   //    publishMsgPayload : Array[0..511] of Byte;
   //    receivedTopic : WString;
   //    receivedMsgPayload : Array[0..1024] of Byte;
   //    valid : Bool;
   //    done : Bool;
   //    busy : Bool;
   //    error : Bool;
   //    status : Word;
   //    diagnostics : "typeDiagnostics";
   //    receivedMsgStatus : USInt;
   //    receivedMsgDataLen : UDInt;
   // END_VAR
BEGIN
END_DATA_BLOCK

DATA_BLOCK "Light_Bars_DB_1"   // DB235
VERSION : 0.1
// stored: AutoNumber true, DBAccessibleFromOPCUA true, InstanceOfName Light_Bars, InstanceOfType FB
"Light_Bars"
BEGIN
END_DATA_BLOCK

DATA_BLOCK "Light_Bars_DB_2"   // DB41
VERSION : 0.1
// stored: AutoNumber true, DBAccessibleFromOPCUA true, InstanceOfName Light_Bars, InstanceOfType FB
"Light_Bars"
BEGIN
END_DATA_BLOCK

DATA_BLOCK "Light_Bars_DB_3"   // DB237
VERSION : 0.1
// stored: AutoNumber true, DBAccessibleFromOPCUA true, InstanceOfName Light_Bars, InstanceOfType FB
"Light_Bars"
BEGIN
END_DATA_BLOCK

DATA_BLOCK "Light_Bars_DB_4"   // DB236
VERSION : 0.1
// stored: AutoNumber true, DBAccessibleFromOPCUA true, InstanceOfName Light_Bars, InstanceOfType FB
"Light_Bars"
BEGIN
END_DATA_BLOCK

DATA_BLOCK "Light_Bars_DB_5"   // DB234
VERSION : 0.1
// stored: AutoNumber true, DBAccessibleFromOPCUA true, InstanceOfName Light_Bars, InstanceOfType FB
"Light_Bars"
BEGIN
END_DATA_BLOCK

DATA_BLOCK "MQTT_Handler_FB_DB"   // DB44
VERSION : 0.1
// stored: AutoNumber true, DBAccessibleFromOPCUA true, InstanceOfName MQTT_Handler_FB, InstanceOfType FB
"MQTT_Handler_FB"
BEGIN
END_DATA_BLOCK

DATA_BLOCK "Main_Panel_DB"   // DB11, F_DB
VERSION : 0.1
// stored: AutoNumber true, DBAccessibleFromOPCUA true, InstanceOfName Main_Panel, InstanceOfType FB
"Main_Panel"
BEGIN
END_DATA_BLOCK

DATA_BLOCK "Main_Safety_RTG1_DB"   // DB7, F_DB
NAME : FUSI
VERSION : 0.1
// stored: AutoNumber true, DBAccessibleFromOPCUA true, InstanceOfName Main_Safety_RTG1, InstanceOfType FB
"Main_Safety_RTG1"
BEGIN
END_DATA_BLOCK

DATA_BLOCK "OPC_Control_FB_DB_1"   // DB17
VERSION : 0.1
// stored: AutoNumber true, DBAccessibleFromOPCUA true, InstanceOfName OPC_Control_FB, InstanceOfType FB
"OPC_Control_FB"
BEGIN
END_DATA_BLOCK

DATA_BLOCK "OPC_Control_FB_DB_2"   // DB335
VERSION : 0.1
// stored: AutoNumber true, DBAccessibleFromOPCUA true, InstanceOfName OPC_Control_FB, InstanceOfType FB
"OPC_Control_FB"
BEGIN
END_DATA_BLOCK

DATA_BLOCK "OPC_Control_FB_DB_3"   // DB332
VERSION : 0.1
// stored: AutoNumber true, DBAccessibleFromOPCUA true, InstanceOfName OPC_Control_FB, InstanceOfType FB
"OPC_Control_FB"
BEGIN
END_DATA_BLOCK

DATA_BLOCK "OPC_Control_FB_DB_4"   // DB334
VERSION : 0.1
// stored: AutoNumber true, DBAccessibleFromOPCUA true, InstanceOfName OPC_Control_FB, InstanceOfType FB
"OPC_Control_FB"
BEGIN
END_DATA_BLOCK

DATA_BLOCK "OPC_Control_FB_DB_5"   // DB333
VERSION : 0.1
// stored: AutoNumber true, DBAccessibleFromOPCUA true, InstanceOfName OPC_Control_FB, InstanceOfType FB
"OPC_Control_FB"
BEGIN
END_DATA_BLOCK

DATA_BLOCK "Order_Table_FB_DB_1"   // DB139
VERSION : 0.1
// stored: AutoNumber true, DBAccessibleFromOPCUA true, InstanceOfName Order_Table_FB, InstanceOfType FB
"Order_Table_FB"
BEGIN
END_DATA_BLOCK

DATA_BLOCK "Order_Table_FB_DB_2"   // DB324
VERSION : 0.1
// stored: AutoNumber true, DBAccessibleFromOPCUA true, InstanceOfName Order_Table_FB, InstanceOfType FB
"Order_Table_FB"
BEGIN
END_DATA_BLOCK

DATA_BLOCK "Order_Table_FB_DB_3"   // DB326
VERSION : 0.1
// stored: AutoNumber true, DBAccessibleFromOPCUA true, InstanceOfName Order_Table_FB, InstanceOfType FB
"Order_Table_FB"
BEGIN
END_DATA_BLOCK

DATA_BLOCK "Order_Table_FB_DB_4"   // DB327
VERSION : 0.1
// stored: AutoNumber true, DBAccessibleFromOPCUA true, InstanceOfName Order_Table_FB, InstanceOfType FB
"Order_Table_FB"
BEGIN
END_DATA_BLOCK

DATA_BLOCK "Order_Table_FB_DB_5"   // DB325
VERSION : 0.1
// stored: AutoNumber true, DBAccessibleFromOPCUA true, InstanceOfName Order_Table_FB, InstanceOfType FB
"Order_Table_FB"
BEGIN
END_DATA_BLOCK

DATA_BLOCK "Remote_Panel_DB_1"   // DB8, F_DB
VERSION : 0.1
// stored: AutoNumber true, DBAccessibleFromOPCUA true, InstanceOfName Remote_Panel, InstanceOfType FB
"Remote_Panel"
BEGIN
END_DATA_BLOCK

DATA_BLOCK "Remote_Panel_DB_2"   // DB10, F_DB
VERSION : 0.1
// stored: AutoNumber true, DBAccessibleFromOPCUA true, InstanceOfName Remote_Panel, InstanceOfType FB
"Remote_Panel"
BEGIN
END_DATA_BLOCK

DATA_BLOCK "Remote_Panel_DB_3"   // DB156, F_DB
VERSION : 0.1
// stored: AutoNumber true, DBAccessibleFromOPCUA true, InstanceOfName Remote_Panel, InstanceOfType FB
"Remote_Panel"
BEGIN
END_DATA_BLOCK

DATA_BLOCK "Remote_Panel_DB_4"   // DB157, F_DB
VERSION : 0.1
// stored: AutoNumber true, DBAccessibleFromOPCUA true, InstanceOfName Remote_Panel, InstanceOfType FB
"Remote_Panel"
BEGIN
END_DATA_BLOCK

DATA_BLOCK "Remote_Panel_DB_5"   // DB154, F_DB
VERSION : 0.1
// stored: AutoNumber true, DBAccessibleFromOPCUA true, InstanceOfName Remote_Panel, InstanceOfType FB
"Remote_Panel"
BEGIN
END_DATA_BLOCK

DATA_BLOCK "SICK_AFx60_DB_1"   // DB121
VERSION : 0.1
// stored: AutoNumber true, DBAccessibleFromOPCUA true, InstanceOfName FB_SICK_AFx60_PN, InstanceOfType FB
"FB_SICK_AFx60_PN"
BEGIN
END_DATA_BLOCK

DATA_BLOCK "SICK_AFx60_DB_2"   // DB319
VERSION : 0.1
// stored: AutoNumber true, DBAccessibleFromOPCUA true, InstanceOfName FB_SICK_AFx60_PN, InstanceOfType FB
"FB_SICK_AFx60_PN"
BEGIN
END_DATA_BLOCK

DATA_BLOCK "SICK_AFx60_DB_3"   // DB317
VERSION : 0.1
// stored: AutoNumber true, DBAccessibleFromOPCUA true, InstanceOfName FB_SICK_AFx60_PN, InstanceOfType FB
"FB_SICK_AFx60_PN"
BEGIN
END_DATA_BLOCK

DATA_BLOCK "SICK_AFx60_DB_4"   // DB316
VERSION : 0.1
// stored: AutoNumber true, DBAccessibleFromOPCUA true, InstanceOfName FB_SICK_AFx60_PN, InstanceOfType FB
"FB_SICK_AFx60_PN"
BEGIN
END_DATA_BLOCK

DATA_BLOCK "SICK_AFx60_DB_5"   // DB318
VERSION : 0.1
// stored: AutoNumber true, DBAccessibleFromOPCUA true, InstanceOfName FB_SICK_AFx60_PN, InstanceOfType FB
"FB_SICK_AFx60_PN"
BEGIN
END_DATA_BLOCK

DATA_BLOCK "SICK_Lector_Control_DB_1"   // DB47
VERSION : 0.1
// stored: AutoNumber true, DBAccessibleFromOPCUA true, InstanceOfName SICK_Lector_Control_FB, InstanceOfType FB
"SICK_Lector_Control_FB"
BEGIN
END_DATA_BLOCK

DATA_BLOCK "SICK_Lector_Control_DB_2"   // DB63
VERSION : 0.1
// stored: AutoNumber true, DBAccessibleFromOPCUA true, InstanceOfName SICK_Lector_Control_FB, InstanceOfType FB
"SICK_Lector_Control_FB"
BEGIN
END_DATA_BLOCK

DATA_BLOCK "SICK_Lector_Control_DB_3"   // DB48
VERSION : 0.1
// stored: AutoNumber true, DBAccessibleFromOPCUA true, InstanceOfName SICK_Lector_Control_FB, InstanceOfType FB
"SICK_Lector_Control_FB"
BEGIN
END_DATA_BLOCK

DATA_BLOCK "SICK_Lector_Control_DB_4"   // DB153
VERSION : 0.1
// stored: AutoNumber true, DBAccessibleFromOPCUA true, InstanceOfName SICK_Lector_Control_FB, InstanceOfType FB
"SICK_Lector_Control_FB"
BEGIN
END_DATA_BLOCK

DATA_BLOCK "SICK_Lector_Control_DB_5"   // DB155
VERSION : 0.1
// stored: AutoNumber true, DBAccessibleFromOPCUA true, InstanceOfName SICK_Lector_Control_FB, InstanceOfType FB
"SICK_Lector_Control_FB"
BEGIN
END_DATA_BLOCK

DATA_BLOCK "SICK_Lector_FB_DB_1"   // DB45
AUTHOR : SICKAG
FAMILY : Ident
VERSION : 1.2
// stored: AutoNumber true, DBAccessibleFromOPCUA true, InstanceOfName SICK_Lector_CLV6xx_PNDP, InstanceOfType FB
"SICK_Lector_CLV6xx_PNDP"
BEGIN
END_DATA_BLOCK

DATA_BLOCK "SICK_Lector_FB_DB_2"   // DB306
AUTHOR : SICKAG
FAMILY : Ident
VERSION : 1.2
// stored: AutoNumber true, DBAccessibleFromOPCUA true, InstanceOfName SICK_Lector_CLV6xx_PNDP, InstanceOfType FB
"SICK_Lector_CLV6xx_PNDP"
BEGIN
END_DATA_BLOCK

DATA_BLOCK "SICK_Lector_FB_DB_3"   // DB74
AUTHOR : SICKAG
FAMILY : Ident
VERSION : 1.2
// stored: AutoNumber true, DBAccessibleFromOPCUA true, InstanceOfName SICK_Lector_CLV6xx_PNDP, InstanceOfType FB
"SICK_Lector_CLV6xx_PNDP"
BEGIN
END_DATA_BLOCK

DATA_BLOCK "SICK_Lector_FB_DB_4"   // DB131
AUTHOR : SICKAG
FAMILY : Ident
VERSION : 1.2
// stored: AutoNumber true, DBAccessibleFromOPCUA true, InstanceOfName SICK_Lector_CLV6xx_PNDP, InstanceOfType FB
"SICK_Lector_CLV6xx_PNDP"
BEGIN
END_DATA_BLOCK

DATA_BLOCK "SICK_Lector_FB_DB_5"   // DB115
AUTHOR : SICKAG
FAMILY : Ident
VERSION : 1.2
// stored: AutoNumber true, DBAccessibleFromOPCUA true, InstanceOfName SICK_Lector_CLV6xx_PNDP, InstanceOfType FB
"SICK_Lector_CLV6xx_PNDP"
BEGIN
END_DATA_BLOCK

DATA_BLOCK "Sf_C1101_FB_DB"   // DB243
VERSION : 0.1
// stored: AutoNumber true, DBAccessibleFromOPCUA true, InstanceOfName Safety_Stops_FB, InstanceOfType FB
"Safety_Stops_FB"
BEGIN
END_DATA_BLOCK

DATA_BLOCK "Sf_C1102_FB_DB"   // DB253
VERSION : 0.1
// stored: AutoNumber true, DBAccessibleFromOPCUA true, InstanceOfName Safety_Stops_FB, InstanceOfType FB
"Safety_Stops_FB"
BEGIN
END_DATA_BLOCK

DATA_BLOCK "Sf_C1103_FB_DB"   // DB250
VERSION : 0.1
// stored: AutoNumber true, DBAccessibleFromOPCUA true, InstanceOfName Safety_Stops_FB, InstanceOfType FB
"Safety_Stops_FB"
BEGIN
END_DATA_BLOCK

DATA_BLOCK "Sf_C1104_FB_DB"   // DB249
VERSION : 0.1
// stored: AutoNumber true, DBAccessibleFromOPCUA true, InstanceOfName Safety_Stops_FB, InstanceOfType FB
"Safety_Stops_FB"
BEGIN
END_DATA_BLOCK

DATA_BLOCK "Sf_C1105_FB_DB"   // DB245
VERSION : 0.1
// stored: AutoNumber true, DBAccessibleFromOPCUA true, InstanceOfName Safety_Stops_FB, InstanceOfType FB
"Safety_Stops_FB"
BEGIN
END_DATA_BLOCK

DATA_BLOCK "Sf_C1106_FB_DB"   // DB246
VERSION : 0.1
// stored: AutoNumber true, DBAccessibleFromOPCUA true, InstanceOfName Safety_Stops_FB, InstanceOfType FB
"Safety_Stops_FB"
BEGIN
END_DATA_BLOCK

DATA_BLOCK "Sf_C1107_FB_DB"   // DB256
VERSION : 0.1
// stored: AutoNumber true, DBAccessibleFromOPCUA true, InstanceOfName Safety_Stops_FB, InstanceOfType FB
"Safety_Stops_FB"
BEGIN
END_DATA_BLOCK

DATA_BLOCK "Sf_C1108_FB_DB"   // DB248
VERSION : 0.1
// stored: AutoNumber true, DBAccessibleFromOPCUA true, InstanceOfName Safety_Stops_FB, InstanceOfType FB
"Safety_Stops_FB"
BEGIN
END_DATA_BLOCK

DATA_BLOCK "Sf_C1201_FB_DB"   // DB247
VERSION : 0.1
// stored: AutoNumber true, DBAccessibleFromOPCUA true, InstanceOfName Safety_Stops_FB, InstanceOfType FB
"Safety_Stops_FB"
BEGIN
END_DATA_BLOCK

